TYPE "UDT_Divert_Constraint_Setting"
VERSION : 0.1
   STRUCT
      Enable : Bool := FALSE;
      Threshold : Int;
      Priority : Int;
      Sort_Code : Int;
      Preferred_Direction : Byte := 16#00;   // Bit0 = Wait Bit1= Straight Bit2= Left Bit3 = Right
      Disallowed_Direction : Byte := 16#00;   // Bit0 = Wait Bit1= Straight Bit2= Left Bit3 = Right
   END_STRUCT;

END_TYPE

TYPE "UDT_SWS_Servo_Setting"
VERSION : 0.1
   STRUCT
      Enable_Soft_Limit { ExternalAccessible := 'False'; ExternalVisible := 'False'; ExternalWritable := 'False'} : Bool := TRUE;
      Enable_Hard_Limit { ExternalAccessible := 'False'; ExternalVisible := 'False'; ExternalWritable := 'False'} : Bool;
      Continuous_Action_Mode : Bool := TRUE;
      STOUsed : Bool;
      Left_Position_Setpoint : Int := -60;   // [°]
      Right_Position_Setpoint : Int := 60;   // [°]
      Speed_Setpoint : Int := 1200;   // [°/s]
      Acc_Setpoint { ExternalAccessible := 'False'; ExternalVisible := 'False'; ExternalWritable := 'False'} : Int := 20000;   // [°/s²]
      Dec_Setpoint { ExternalAccessible := 'False'; ExternalVisible := 'False'; ExternalWritable := 'False'} : Int := 20000;   // [°/s²]
      Max_Left_Position { ExternalAccessible := 'False'; ExternalVisible := 'False'; ExternalWritable := 'False'} : Int := -65;   // [°]
      Max_Right_Position { ExternalAccessible := 'False'; ExternalVisible := 'False'; ExternalWritable := 'False'} : Int := 65;   // [°]
      Max_Speed { ExternalAccessible := 'False'; ExternalVisible := 'False'; ExternalWritable := 'False'} : Int := 1500;   // [°/s]
   END_STRUCT;

END_TYPE

TYPE "UDT_SWS_Roller_Hardware_Setting"
VERSION : 0.1
   STRUCT
      Module_Roller_Count : Int := 29;
      Speed_Straight : Int := 1200;
      Speed_Left : Int := 1500;
      Speed_Right : Int := 1500;
      Reference_RPM : Real := 470.0;
      Acceleration : Int := 4000;   // [mm/s²] Ramp up
      Deceleration : Int := 4000;   // [mm/s²] Ramp down
   END_STRUCT;

END_TYPE

TYPE "i_udtSettings"
VERSION : 0.1
   STRUCT
      timStartReadDelay : UDInt := 40;   // Start read delay time (mseconds)
      timSpare_Timer2 : UDInt;   // Not in use
      timNoActivity : UDInt := 10000;   // Time to consider Camera not working ok
      timTimeOutRead : UDInt := 400;   // TimeOut to get Barcode (mseconds)
      TimeStarting : UDInt := 5000;   // Time starting camera (waitting for normal operation)
      timTrshNoReadRow : Int;   // threshold no reads in a row
      xIndexProtocol : Bool := TRUE;   // 1: In Use; 0: Not used
      xIOConditioning : Bool := FALSE;   // 1: In Use; 0: Not used
      xFocusingDevice : Bool := FALSE;
      Protocol : Struct
         Encapsulation : Bool := TRUE;
         Header : String := '$02';
         Footer : String := '$03';
         Separator : String := '€';
         VirtualID : String := '!';
         ValidTelegram : String := '*';
         NoRead : String := '??????????';
         MultiRead : String := '9999999999';
      END_STRUCT;
      Telegrams : Struct
         Number : Int := 4;
         Parameters : Array[0..10] of Struct
            Length : Int;   // Telegram length without encapsulation
            "Type" : Int;   // 0: No Code; 1: Status Telegram; 2: Barcode Telegram; 9: Special Barcode Telegram
            ID : Char;   // Telegram ID. D: Status; I: Index Barcode
            Barcode : Struct   // Only for Types > 2
               FromDAD : String;
               ToPLC : String := '0000000000';
            END_STRUCT;
         END_STRUCT;
      END_STRUCT;
   END_STRUCT;

END_TYPE

TYPE "UDT_G115D_Setting"
VERSION : 0.1
   STRUCT
      Speed1 : Int := 1000;   // [mm/s] Target speed 1
      Speed2 : Int := 500;   // [mm/s] Target speed 2
      Speed3 : Int;   // [mm/s] Target speed 3
      Speed4 : Int;   // [mm/s] Target speed 4
      Acceleration : Int := 4000;   // [mm/s²] Ramp up
      Deceleration : Int := 4000;   // [mm/s²] Ramp down
      RefSpeed : Int;   // [mm/s] Speed at 3000RPM
      RefRampTime : Int := 10000;   // [ms] Ramp up and ramp down time for 3000RPM
      Magnetization_Delay : Int;   // [ms] Delay time from run command to mote have speed
      ReverseDirection : Bool;   // TRUE = Reverse inverter output direction
      STOUsed : Bool;   // TRUE = STO is used
   END_STRUCT;

END_TYPE

TYPE "UDT_MultiControl_HW_Diagnostics"
VERSION : 0.1
   STRUCT
      RD1_Run_Command : Bool;   // Rum command from controller
      RD2_Run_Command : Bool;   // Rum command from controller
      RD3_Run_Command : Bool;   // Rum command from controller
      RD4_Run_Command : Bool;   // Rum command from controller
      RD1_Actual_Speed : Int;   // [mm/s] Motor actual speed
      RD2_Actual_Speed : Int;   // [mm/s] Motor actual speed
      RD3_Actual_Speed : Int;   // [mm/s] Motor actual speed
      RD4_Actual_Speed : Int;   // [mm/s] Motor actual speed
      Control_Voltage : Int;   // [mV] Control logic voltage
      Motor_Voltage : Int;   // [mV] Motor voltage
      Temperature : Int;   // [0,1°] Temperature
      RD1_Actual_Current : Int;   // [mA] Actual current
      RD2_Actual_Current : Int;   // [mA] Actual current
      RD3_Actual_Current : Int;   // [mA] Actual current
      RD4_Actual_Current : Int;   // [mA] Actual current
      Motor_Start_Stop_Count : UInt;   // Count of motor start and stop
      Motor_Direction_Switch_Count : UInt;   // Count of motor switch direction
      Motor_Started_Time : UDInt;   // [s] Count time of motor running
   END_STRUCT;

END_TYPE

TYPE "UDT_PEC_Position_Setting"
TITLE = UDT_Sett_PEC
VERSION : 0.1
//Setting of photo electric cell
//# Block Info
//- Title:            UDT_Sett_PEC
//- Comment/Function: Setting of photo electric cell
//- Library/Family:   APS
//- Author:           Jay Liu
//- Tested with:      ---
//- Engineering:      TIA Portal V20
//- Restrictions:     ---
//- Requirements:     ---
//
//# History
// |Version  | Date       | Author                 | Description                   |
// |---------|------------|------------------------|------------------------------ |
// |01.00.00 | 2026-01-22 | Jay Liu                | First released version        |
   STRUCT
      Blockage_Length : DInt := 3000;   // [mm] Delay for detecting a PEC blockage during the running
      Delay_On : DInt := 50;   // [mm] Delay on leading edge of product (flap filter)
      Delay_Off : DInt := 50;   // [mm] Delay off trailing edge of product (flap filter)
      Shifting_Offset : DInt;   // [mm] Shift offset of PE signal
      Handover_Offset : DInt;   // [mm] Distance between PE and the end of section
      Detect_PEC_OnStopped : Bool := TRUE;   // TRUE = Enable delay timer even the section is not running
      Reset_Block_PEC_Oc : Bool;   // TRUE = Allow reset of blockage error with PEC still covered
      Item_On : Bool;   // TRUE = When detect item the input signal should be true FALSE= When detect item the input signal should be false
   END_STRUCT;

END_TYPE

TYPE "UDT_TCON_PAR"
VERSION : 0.1
   STRUCT
      InterfaceId : HW_ANY := 64;
      ID : CONN_OUC := 1;
      ConnectionType : Byte := 11;
      ActiveEstablished : Bool;
      RemoteAddress {InstructionName := 'IP_V4'; LibVersion := '1.0'} : IP_V4;
      RemotePort : UInt;
      LocalPort : UInt := 6000;
   END_STRUCT;

END_TYPE

TYPE "UDT_Divert_Decision_Setting"
VERSION : 0.1
   STRUCT
      Decision_Position : DInt;
      Straight_Destination { S7_SetPoint := 'True'} : Int;
      Left_Destination { S7_SetPoint := 'True'} : Int;
      Right_Destination { S7_SetPoint := 'True'} : Int;
      High_Priority { S7_SetPoint := 'True'} : Int := 2;   // Bit0 = Wait Bit1= Straight Bit2= Left Bit3 = Right
      Middle_Priority { S7_SetPoint := 'True'} : Int := 4;   // Bit0 = Wait Bit1= Straight Bit2= Left Bit3 = Right
      Low_Priority { S7_SetPoint := 'True'} : Int := 8;   // Bit0 = Wait Bit1= Straight Bit2= Left Bit3 = Right
      Default_Direction : Int := 8;   // Bit0 = Wait Bit1= Straight Bit2= Left Bit3 = Right
      Allow_Wait : Bool := FALSE;
      Destination_Invalid : "UDT_Divert_Constraint_Setting" := ((), (), 1, 7, (), ());
      No_Destination : "UDT_Divert_Constraint_Setting" := ((), (), 2, 16, (), ());
      Gap_Error : "UDT_Divert_Constraint_Setting" := ((), 250, 4, 4, (), ());
      Diemension_Error : "UDT_Divert_Constraint_Setting" := ((), 700, 6, 18, (), ());
      Throughput_Limit_Straight : "UDT_Divert_Constraint_Setting" := ((), (), 10, 13, (), ());
      Throughput_Limit_Left : "UDT_Divert_Constraint_Setting" := ((), (), 10, 13, (), ());
      Throughput_Limit_Right : "UDT_Divert_Constraint_Setting" := ((), (), 10, 13, (), ());
      Dir_Fault_Straight : "UDT_Divert_Constraint_Setting" := ((), (), 13, 20, (), ());
      Dir_Fault_Left : "UDT_Divert_Constraint_Setting" := ((), (), 13, 20, (), ());
      Dir_Fault_Right : "UDT_Divert_Constraint_Setting" := ((), (), 13, 20, (), ());
      Dir_Disabled_Straight : "UDT_Divert_Constraint_Setting" := ((), (), 14, 12, (), ());
      Dir_Disabled_Left : "UDT_Divert_Constraint_Setting" := ((), (), 14, 12, (), ());
      Dir_Disabled_Right : "UDT_Divert_Constraint_Setting" := ((), (), 14, 12, (), ());
      Dir_Full_Straight : "UDT_Divert_Constraint_Setting" := ((), (), 15, 5, (), ());
      Dir_Full_Left : "UDT_Divert_Constraint_Setting" := ((), (), 15, 5, (), ());
      Dir_Full_Right : "UDT_Divert_Constraint_Setting" := ((), (), 15, 5, (), ());
      No_Read : "UDT_Divert_Constraint_Setting" := ((), (), 16, 8, (), ());
      No_Code : "UDT_Divert_Constraint_Setting" := ((), (), 17, 9, (), ());
      Multi_Read : "UDT_Divert_Constraint_Setting" := ((), (), 18, 10, (), ());
      Unexpected_Item : "UDT_Divert_Constraint_Setting" := ((), (), 19, 2, (), ());
   END_STRUCT;

END_TYPE

TYPE "UDT_SWS_Divert_Setting"
VERSION : 0.1
   STRUCT
      Fixed_Ratio_Staight : Int;
      Fixed_Ratio_Left : Int;
      Fixed_Ratio_Right : Int;
      First_Group_Action_Delay : Int := 350;
      Group2_Action_Delay : Int := 160;
      Group3_Action_Delay : Int := 160;
      Group4_Action_Delay : Int := 160;
      Group5_Action_Delay : Int := 160;
      Group6_Action_Delay : Int := 160;
      Group7_Action_Delay : Int := 160;
      Group8_Action_Delay : Int := 160;
      Group9_Action_Delay : Int := 160;
   END_STRUCT;

END_TYPE

TYPE "UDT_SWS_Hardware_Setting"
VERSION : 0.1
   STRUCT
      Roller { S7_SetPoint := 'False'} : "UDT_SWS_Roller_Hardware_Setting" := (29, 1200, 1500, 1500, 470.0, 4000, 4000);
      Servo_U401 : "UDT_SWS_Servo_Setting" := ((), (), (), (), -30, 30, (), (), (), (), (), ());
      Servo_U411 : "UDT_SWS_Servo_Setting" := ((), (), (), (), -45, 45, (), (), (), (), (), ());
      Servo_U421 : "UDT_SWS_Servo_Setting";
      Servo_U431 : "UDT_SWS_Servo_Setting";
      Servo_U441 : "UDT_SWS_Servo_Setting";
      Servo_U451 : "UDT_SWS_Servo_Setting";
      Servo_U461 : "UDT_SWS_Servo_Setting";
      Servo_U471 : "UDT_SWS_Servo_Setting";
      Servo_U481 : "UDT_SWS_Servo_Setting";
   END_STRUCT;

END_TYPE

TYPE "UDT_MultiControl_Setting"
VERSION : 0.1
   STRUCT
      Speed1 : Int := 1000;   // [mm/s] Target speed 1
      Speed2 : Int := 500;   // [mm/s] Target speed 2
      Speed3 : Int;   // [mm/s] Target speed 3
      Speed4 : Int;   // [mm/s] Target speed 4
      Acceleration : Int := 4000;   // [mm/s²] Ramp up
      Deceleration : Int := 4000;   // [mm/s²] Ramp down
      RefSpeed : Int := 1390;   // [mm/s] Reference Speed
      RD1_Motor_Number : Int;
      RD2_Motor_Number : Int;
      RD3_Motor_Number : Int;
      RD4_Motor_Number : Int;
      ReverseDirection : Bool;
   END_STRUCT;

END_TYPE

TYPE "UDT_G115D_HW_Diagnostics"
VERSION : 0.1
   STRUCT
      Run_Command : Bool;   // Rum command from controller
      Brake_Open : Bool;   // Holding brake open
      DI0 : Bool;   // Digital input 0 status
      DI1 : Bool;   // Digital input 1 status
      DI2 : Bool;   // Digital input 2 status
      DI3 : Bool;   // Digital input 3 status
      DIO24 : Bool;   // Digital input/output 24 status
      DIO25 : Bool;   // Digital input/output 25 status
      Memory_Card_In : Bool;   // Memory card is inserted
      Memory_Card_Active : Bool;   // Memory card is active
      PN_Port1_Down : Bool;   // Profinet port 1 up
      PN_Port2_Down : Bool;   // Profinet port 2 up
      Actual_Speed : Int;   // [mm/s] Motor Actual Speed
      DCLink_Voltage : Int;   // [V] DC link voltage
      Actual_Current : Int;   // [0.1A] Actual current
      Active_Power : Int;   // [W] Active power
      Motor_Start_Stop_Count : UInt;   // Count of motor start and stop
      Motor_Direction_Switch_Count : UInt;   // Count of motor switch direction
      Motor_Started_Time : UDInt;   // [s] Count time of motor running
   END_STRUCT;

END_TYPE

TYPE "UDT_SWS_Roller_Interface_Setting"
VERSION : 0.1
   STRUCT
      Status_Interval : Time := T#200ms;
      Num_Of_Comm_Error : Int := 3;
   END_STRUCT;

END_TYPE

TYPE "UDT_G115D_HW_Input"
VERSION : 0.1
   STRUCT
      ZSW1_Bit00_ReadyOn : Bool;   // 0: Ready for switching on
      ZSW1_Bit01_Ready : Bool;   // 1: Ready (operating condition)
      ZSW1_Bit02_Enabled : Bool;   // 2: Operation enabled
      ZSW1_Bit03_Fault : Bool;   // 3: Fault present (1: fault)
      ZSW1_Bit04_NoCoastActive : Bool;   // 4: No coast down active (0: active)
      ZSW1_Bit05_NoQuickStopActive : Bool;   // 5: No quick stop active (0: active)
      ZSW1_Bit06_Inhibit : Bool;   // 6: Switching on inhibited
      ZSW1_Bit07_Alarm : Bool;   // 7: Alarm present (1: alarm)
      ZSW1_Bit08_DeviationOK : Bool;   // 8: Setpoint/actual value deviation
      ZSW1_Bit09_ControlQuest : Bool;   // 9: Control requested
      ZSW1_Bit10_OverSpeed : Bool;   // 10: f or n comparison value reached
      ZSW1_Bit11_Limit : Bool;   // 11: Torque limit not reached
      ZSW1_Bit12_Brake : Bool;   // 12: Holding brake open
      ZSW1_Bit13_MotorTempOK : Bool;   // 13: Motor temperature OK (1: OK)
      ZSW1_Bit14_Direction_CW : Bool;   // 14: n_act >= 0 (1: positive)
      ZSW1_Bit15_VFDTempOK : Bool;   // 15: Reserved Speed actual value (NIST_A)
      NIST_A : Int;   // Actual speed (-16384 to +16384)
      ZSW_G115D_Bit00_DI0 : Bool;   // 0: Digital input 0 status
      ZSW_G115D_Bit01_DI1 : Bool;   // 1: Digital input 1 status
      ZSW_G115D_Bit02_DI2 : Bool;   // 2: Digital input 2 status
      ZSW_G115D_Bit03_DI3 : Bool;   // 3: Digital input 3 status
      ZSW_G115D_Bit04_DIO24 : Bool;   // 4: DI/O 24 status
      ZSW_G115D_Bit05_DIO25 : Bool;   // 5: DI/O 25 status
      ZSW_G115D_Bit06_STOActive : Bool;   // 6: STO is active
      ZSW_G115D_Bit07_Reserved : Bool;   // 7: Reserved
      ZSW_G115D_Bit08_PowerOff : Bool;   // 8: Power switch OFF status
      ZSW_G115D_Bit09_Auto : Bool;   // 9: Automatic mode active
      ZSW_G115D_Bit10_Manual : Bool;   // 10: Manual mode active
      ZSW_G115D_Bit11_Bypass : Bool;   // 11: Stop/Slow bypass activated
      ZSW_G115D_Bit12_ContMotion : Bool;   // 12: Continuous motion activated
      ZSW_G115D_Bit13_JogLeft : Bool;   // 13: Motor jogging to the left
      ZSW_G115D_Bit14_JogRight : Bool;   // 14: Motor jogging to the right
      ZSW_G115D_Bit15_Reserved : Bool;   // 15: Reserved Fault and alarm codes
      FaultCode : Word;   // Fault code (0: no fault)
      AlarmCode : Word;   // Alarm code (0: no alarm)
      DCLinkVoltage : Int;   // DC link voltage [V]
      ActualCurrent : Int;   // Actual current [0.1A]
      ActivePower : Int;   // Active power [W]
      ZSW2_G115D_Bit00_Memory_Card_In : Bool;
      ZSW2_G115D_Bit01_Memory_Card_Active : Bool;
      ZSW2_G115D_Bit02_Memory_Card_Siemens : Bool;
      ZSW2_G115D_Bit03_Memory_Card_USB : Bool;
      ZSW2_G115D_Bit04_Reserved : Bool;
      ZSW2_G115D_Bit05_Reserved : Bool;
      ZSW2_G115D_Bit06_Reserved : Bool;
      ZSW2_G115D_Bit07_Reserved : Bool;
      ZSW2_G115D_Bit08_Reserved : Bool;
      ZSW2_G115D_Bit09_Reserved : Bool;
      ZSW2_G115D_Bit10_Reserved : Bool;
      ZSW2_G115D_Bit11_Reserved : Bool;
      ZSW2_G115D_Bit12_Reserved : Bool;
      ZSW2_G115D_Bit13_Reserved : Bool;
      ZSW2_G115D_Bit14_Reserved : Bool;
      ZSW2_G115D_Bit15_Reserved : Bool;
   END_STRUCT;

END_TYPE

TYPE "UDT_S210_Speed_Setting"
VERSION : 0.1
   STRUCT
      Speed1 : Int := 1000;   // [mm/s] Target speed 1
      Speed2 : Int := 500;   // [mm/s] Target speed 2
      Speed3 : Int;   // [mm/s] Target speed 3
      Speed4 : Int;   // [mm/s] Target speed 4
      Acceleration : Int := 4000;   // [mm/s²] Ramp up
      Deceleration : Int := 4000;   // [mm/s²] Ramp down
      MinSpeed : Int := 500;   // [mm/s] Minimum target speed
      MaxSpeed : Int := 2500;   // [mm/s] Maximum target speed
      Continuous_Action_Mode : Bool := TRUE;
      Use_Hardware_Feedback : Bool;
      ReverseDirection : Bool;
      STOUsed : Bool;
   END_STRUCT;

END_TYPE

TYPE "UDT_G115D_HW_Output"
VERSION : 0.1
   STRUCT
      STW1_Bit00_On : Bool;   // 0: ON/OFF1 command (0->1: ON)
      STW1_Bit01_Off2 : Bool;   // 1: No OFF2 command (0: active, coast stop)
      STW1_Bit02_Off3 : Bool;   // 2: No OFF3 command (0: active, quick stop)
      STW1_Bit03_Enable : Bool;   // 3: Operation enable
      STW1_Bit04_RampEnable : Bool;   // 4: Ramp-function generator enable
      STW1_Bit05_RampContinue : Bool;   // 5: Continue ramp-function generator
      STW1_Bit06_SetEnable : Bool;   // 6: Setpoint enable
      STW1_Bit07_Ack : Bool;   // 7: Acknowledge faults (0->1: acknowledge)
      STW1_Bit08_Reserved : Bool;   // 8: Reserved
      STW1_Bit09_Reserved : Bool;   // 9: Reserved
      STW1_Bit10_PLC : Bool;   // 10: Control by PLC (must be 1)
      STW1_Bit11_Reverse : Bool;   // 11: Reverse (1: reverse direction)
      STW1_Bit12_Reserved : Bool;   // 12: Reserved
      STW1_Bit13_MOP_Up : Bool;   // 13: Motorized potentiometer, raise
      STW1_Bit14_MOP_Down : Bool;   // 14: Motorized potentiometer, lower
      STW1_Bit15_Reserved : Bool;   // 15: Reserved Speed setpoint (NSOLL_A)
      NSOLL_A : Int;   // Speed setpoint (-16384 to +16384)
      STW_G115D_Bit00_DO24 : Bool;   // 0: DO 24 control
      STW_G115D_Bit01_DO25 : Bool;   // 1: DO 25 control
      STW_G115D_Bit02_Disable_StopSlow_Sensor : Bool;   // 2: Stop-Slow bypass
      STW_G115D_Bit03_Reserved : Bool;   // 3: Reserved
      STW_G115D_Bit04_Reserved : Bool;   // 4: Reserved
      STW_G115D_Bit05_Reserved : Bool;   // 5: Reserved
      STW_G115D_Bit06_Reserved : Bool;   // 6: Reserved
      STW_G115D_Bit07_Reserved : Bool;   // 7: Reserved
      STW_G115D_Bit08_Reserved : Bool;   // 8: Reserved
      STW_G115D_Bit09_Reserved : Bool;   // 9: Reserved
      STW_G115D_Bit10_Reserved : Bool;   // 10: Reserved
      STW_G115D_Bit11_Reserved : Bool;   // 11: Reserved
      STW_G115D_Bit12_Reserved : Bool;   // 12: Reserved
      STW_G115D_Bit13_Reserved : Bool;   // 13: Reserved
      STW_G115D_Bit14_Reserved : Bool;   // 14: Reserved
      STW_G115D_Bit15_Reserved : Bool;   // 15: Reserved
      RampUpScaling : Int;   // Ramp-up time scaling (0-200% = 0-32767)
      RampDownScaling : Int;   // Ramp-down time scaling (0-200% = 0-32767)
   END_STRUCT;

END_TYPE

TYPE "UDT_S210_HW_Diagnostics"
VERSION : 0.1
   STRUCT
      Run_Command : Bool;   // Rum command from controller
      DI0 : Bool;   // Digital input 0 status
      DI1 : Bool;   // Digital input 1 status
      DI2 : Bool;   // Digital input 2 status
      DI3 : Bool;   // Digital input 3 status
      DI4 : Bool;   // Digital input 4 status
      PN_Port1_Down : Bool;   // Profinet port 1 up
      PN_Port2_Down : Bool;   // Profinet port 2 up
      Actual_Speed : Int;   // [mm/s] Motor actual speed
      Actual_Displacement : Int;   // [mm/scan] Motor movement distance
      Actual_Position : Real;   // [°] Motor actual position
      DCLink_Voltage : Int;   // [V] DC link voltage
      Actual_Current : Int;   // [0.1A] Actual current
      Active_Power : Int;   // [W] Active power
      Motor_Start_Stop_Count : UInt;   // Count of motor start and stop
      Motor_Direction_Switch_Count : UInt;   // Count of motor switch direction
      Motor_Started_Time : UDInt;   // [s] Count time of motor running
   END_STRUCT;

END_TYPE

TYPE "UDT_Base_Conveyor_Setting"
TITLE = UDT_Sett_Base_Conveyor
VERSION : 0.1
//Setting of base tranpsort control
//# Block Info
//- Title:            UDT_Sett_Base_Conveyor
//- Comment/Function: Setting of base tranpsort control
//- Library/Family:   APS
//- Author:           Jay Liu
//- Tested with:      ---
//- Engineering:      TIA Portal V20
//- Restrictions:     ---
//- Requirements:     ---
//
//# History
// |Version  | Date       | Author                 | Description                   |
// |---------|------------|------------------------|------------------------------ |
// |01.00.00 | 2026-01-22 | Jay Liu                | First released version        |
   STRUCT
      Delay_Dieback : DInt := 50;   // [mm] Delay from end to stop in dieback
      Delay_Startup : DInt := 100;   // [mm] Delay restart after dieback
      Delay_Waiting_Item : DInt;   // [mm] Delay for receive item from upstream
      Delay_Finish_Handover : DInt;   // [mm] Delay handover after items exit the END PEC
      Delay_Energysave : DInt := 5000;   // [mm] Delay running after clearing
      Delay_Cascade_Startup : DInt := 100;   // [mm] Cascade delay 0: Startup immediately
      Delay_Cascade_Shutdown : DInt := -1;   // [ms] Cascade delay -1: disable function 0: Shutdown immediately
      Slave_Mode : Bool;   // TRUE = Make this section a slave
      Enable_DieForward : Bool;   // TRUE = Halt conveyor if upstream handover occurs error
   END_STRUCT;

END_TYPE

TYPE "UDT_Flow_Control_Setting"
TITLE = UDT_Sett_Flow_Control
VERSION : 0.1
//Setting of flow control
//# Block Info
//- Title:            UDT_Sett_Flow_Control
//- Comment/Function: Setting of flow control
//- Library/Family:   APS
//- Author:           Jay Liu
//- Tested with:      ---
//- Engineering:      TIA Portal V20
//- Restrictions:     ---
//- Requirements:     ---
//
//# History
// |Version  | Date       | Author                 | Description                   |
// |---------|------------|------------------------|------------------------------ |
// |01.00.00 | 2026-01-22 | Jay Liu                | First released version        |
   STRUCT
      Minimum_Gap : Int;   // [mm] Minimum gap length between products (0 = no gap control)
      Add_Gap_Stop : Int;   // [mm] Additional gap after stop of upstream conveyor
      Minimum_Head_To_Head : Int;   // [mm] Minimum head to head length (0 = no head to head control)
      Add_Head_To_Head_Stop : Int;   // [mm] Additional head to head length after stop of upstream conveyor
   END_STRUCT;

END_TYPE

TYPE "UDT_PEC_Trigger_Setting"
TITLE = UDT_Sett_PEC
VERSION : 0.1
//Setting of photo electric cell
//# Block Info
//- Title:            UDT_Sett_PEC
//- Comment/Function: Setting of photo electric cell
//- Library/Family:   APS
//- Author:           Jay Liu
//- Tested with:      ---
//- Engineering:      TIA Portal V20
//- Restrictions:     ---
//- Requirements:     ---
//
//# History
// |Version  | Date       | Author                 | Description                   |
// |---------|------------|------------------------|------------------------------ |
// |01.00.00 | 2026-01-22 | Jay Liu                | First released version        |
   STRUCT
      Blockage_Length : Int := 3000;   // [mm] Delay for detecting a PEC blockage during the running
      Delay_On : Int := 50;   // [mm] Delay on leading edge of product (flap filter)
      Delay_Off : Int := 50;   // [mm] Delay off trailing edge of product (flap filter)
      Detect_PEC_OnStopped : Bool := TRUE;   // TRUE = Enable delay timer even the section is not running
      Reset_Block_PEC_Oc : Bool;   // TRUE = Allow reset of blockage error with PEC still covered
      Item_On : Bool;   // TRUE = When detect item the input signal should be true FALSE= When detect item the input signal should be false
   END_STRUCT;

END_TYPE

TYPE "UDT_Track_Statistics"
VERSION : 0.1
   STRUCT
      Last_Slip : Int;
      Last_Data : Int;
      Average_Slip : Real;
      Update_Performance : Real;
      Missing_Items : UDInt;
      UFO_Generated : UDInt;
      Number_Of_Items : UDInt;
   END_STRUCT;

END_TYPE

TYPE "UDT_Mesasuring_Point_Statistics"
VERSION : 0.1
   STRUCT
      Capacity : Int;
      Length : UDInt;
      Window : UDInt;
      Gap : UDInt;
   END_STRUCT;

END_TYPE

TYPE "UDT_Scanner_Statistics"
VERSION : 0.1
   STRUCT
      Total : UDInt;
      GoodRead : UDInt;
      NoRead : UDInt;
      MultiRead : UDInt;
      NoCode : UDInt;
      NoFoundID : UDInt;
      NotDefined : UDInt;
   END_STRUCT;

END_TYPE

TYPE "UDT_Chute_Statistics"
VERSION : 0.1
   STRUCT
      PE_Full_Items : UDInt;
   END_STRUCT;

END_TYPE

TYPE "UDT_IODevice_Diag"
TITLE = UDT_Diag_HW
VERSION : 0.1
//Diagnose data of IO Device
//# Block Info
//- Title:            UDT_Diag_HW
//- Comment/Function: Diagnose data of IO Device
//- Library/Family:   APS
//- Author:           Jay Liu
//- Tested with:      ---
//- Engineering:      TIA Portal V20
//- Restrictions:     ---
//- Requirements:     ---
//
//# History
// |Version  | Date       | Author                 | Description                   |
// |---------|------------|------------------------|------------------------------ |
// |01.00.00 | 2026-01-22 | Jay Liu                | First released version        |
   STRUCT
      Module_Not_Present : Array[0..127] of Bool;   // Module not present
      Module_Error : Array[0..127] of Bool;   // Module error
   END_STRUCT;

END_TYPE

TYPE "UDT_PNIO_System_Diag"
TITLE = UDT_Diag_PNIO_System
VERSION : 0.1
//Diagnose data of IO System
//# Block Info
//- Title:            UDT_Diag_PNIO_System
//- Comment/Function: Diagnose data of IO System
//- Library/Family:   APS
//- Author:           Jay Liu
//- Tested with:      ---
//- Engineering:      TIA Portal V20
//- Restrictions:     ---
//- Requirements:     ---
//
//# History
// |Version  | Date       | Author                 | Description                   |
// |---------|------------|------------------------|------------------------------ |
// |01.00.00 | 2026-01-22 | Jay Liu                | First released version        |
   STRUCT
      Device_Not_Present : Array[0..1023] of Bool;   // Profinet device not present
      Device_Error : Array[0..1023] of Bool;   // Profinet device error
   END_STRUCT;

END_TYPE

TYPE "UDT_Divert_Statistics"
VERSION : 0.1
   STRUCT
      Direction_Straight : UDInt;
      Direction_Left : UDInt;
      Direction_Right : UDInt;
   END_STRUCT;

END_TYPE

TYPE "UDT_G115D_HW_Interface"
VERSION : 0.1
   STRUCT
      Input { S7_SetPoint := 'False'} : "UDT_G115D_HW_Input";
      Output : "UDT_G115D_HW_Output";
   END_STRUCT;

END_TYPE

TYPE "UDT_Conv_Multiple_S210_Diagnostics"
VERSION : 0.1
   STRUCT
      RTS : Bool;   // Section ready to send item
      TIP : Bool;   // Section transfer in porgress
      Downstream_RTR : Bool;   // Downstream section ready to receive item
      Items_Count : UDInt;   // Count of items passed
      Displacement : Int;   // [mm/scan] Conveyor movement distance
      Hardware_U01 { S7_SetPoint := 'False'} : "UDT_S210_HW_Diagnostics";
      Hardware_U02 : "UDT_S210_HW_Diagnostics";
      Hardware_U03 : "UDT_S210_HW_Diagnostics";
      Hardware_U04 : "UDT_S210_HW_Diagnostics";
      Hardware_U05 : "UDT_S210_HW_Diagnostics";
      Hardware_U06 : "UDT_S210_HW_Diagnostics";
      Hardware_U07 : "UDT_S210_HW_Diagnostics";
      Hardware_U08 : "UDT_S210_HW_Diagnostics";
      Hardware_U09 : "UDT_S210_HW_Diagnostics";
      Hardware_U10 : "UDT_S210_HW_Diagnostics";
   END_STRUCT;

END_TYPE

TYPE "UDT_Conv_Dual_G115D_Diagnostics"
VERSION : 0.1
   STRUCT
      RTS : Bool;   // Section ready to send item
      TIP : Bool;   // Section transfer in porgress
      Downstream_RTR : Bool;   // Downstream section ready to receive item
      Items_Count : UDInt;   // Count of items passed
      Displacement : Int;   // [mm/scan] Conveyor movement distance
      Hardware_U01 { S7_SetPoint := 'False'} : "UDT_G115D_HW_Diagnostics";   // Invert driver
      Hardware_U02 : "UDT_G115D_HW_Diagnostics";
   END_STRUCT;

END_TYPE

TYPE "UDT_Conv_Triple_G115D_Diagnostics"
VERSION : 0.1
   STRUCT
      RTS : Bool;   // Section ready to send item
      TIP : Bool;   // Section transfer in porgress
      Downstream_RTR : Bool;   // Downstream section ready to receive item
      Items_Count : UDInt;   // Count of items passed
      Displacement : Int;   // [mm/scan] Conveyor movement distance
      Hardware_U01 { S7_SetPoint := 'False'} : "UDT_G115D_HW_Diagnostics";   // Invert driver
      Hardware_U02 : "UDT_G115D_HW_Diagnostics";
      Hardware_U03 : "UDT_G115D_HW_Diagnostics";
   END_STRUCT;

END_TYPE

TYPE "UDT_Conv_MultiControl_Diagnostics"
VERSION : 0.1
   STRUCT
      RTS : Bool;   // Section ready to send item
      TIP : Bool;   // Section transfer in porgress
      Downstream_RTR : Bool;   // Downstream section ready to receive item
      Items_Count : UDInt;   // Count of items passed
      Displacement : Int;   // [mm/scan] Conveyor movement distance
      Hardware_U01 { S7_SetPoint := 'False'} : "UDT_MultiControl_HW_Diagnostics";   // Invert driver
      Hardware_U02 : "UDT_MultiControl_HW_Diagnostics";
      Hardware_U03 : "UDT_MultiControl_HW_Diagnostics";
      Hardware_U04 : "UDT_MultiControl_HW_Diagnostics";
   END_STRUCT;

END_TYPE

TYPE "UDT_Conv_G115D_Diagnostics"
VERSION : 0.1
   STRUCT
      RTS : Bool;   // Section ready to send item
      TIP : Bool;   // Section transfer in porgress
      Downstream_RTR : Bool;   // Downstream section ready to receive item
      Items_Count : UDInt;   // Count of items passed
      Displacement : Int;   // [mm/scan] Conveyor movement distance
      Hardware { S7_SetPoint := 'False'} : "UDT_G115D_HW_Diagnostics";   // Invert driver
   END_STRUCT;

END_TYPE

TYPE "UDT_MultiControl_HW_Input"
VERSION : 0.1
   STRUCT
      Sensor1 : Bool;
      Sensor2 : Bool;
      Sensor3 : Bool;
      Sensor4 : Bool;
      Sensor5 : Bool;
      Sensor6 : Bool;
      Sensor7 : Bool;
      Sensor8 : Bool;
      Digital_Input_1 : Bool;
      Digital_Input_2 : Bool;
      Digital_Input_3 : Bool;
      Digital_Input_4 : Bool;
      Digital_Input_Spare_1 : Bool;
      Digital_Input_Spare_2 : Bool;
      Digital_Input_Spare_3 : Bool;
      Digital_Input_Spare_4 : Bool;
      MotorErr_RD1 : Bool;
      MotorErr_RD2 : Bool;
      MotorErr_RD3 : Bool;
      MotorErr_RD4 : Bool;
      MotorSpeed_RD1 : SInt;
      MotorSpeed_RD2 : SInt;
      MotorSpeed_RD3 : SInt;
      MotorSpeed_RD4 : SInt;
      MotorStates_Spare : Byte;
      MotorCurrent_RD1 : Int;   // [mA]
      MotorCurrent_RD2 : Int;   // [mA]
      MotorCurrent_RD3 : Int;   // [mA]
      MotorCurrent_RD4 : Int;   // [mA]
      Voltage_Motor : Int;   // [mV]
      Voltage_Control : Int;   // [mV]
      Temperature : Int;   // [0.1C]
      SystemUpTime : UDInt;   // [s]
   END_STRUCT;

END_TYPE

TYPE "UDT_Merge_Singulator_Setting"
VERSION : 0.1
   STRUCT
      StartUp_Delay : Int;   // [ms]
      Dieback_Delay : Int;   // [ms]
   END_STRUCT;

END_TYPE

TYPE "UDT_Echelon_Setting"
VERSION : 0.1
   STRUCT
      StartUp_Delay : Int;   // [ms]
      Dieback_Delay : Int;   // [ms]
   END_STRUCT;

END_TYPE

TYPE "UDT_Tipper_Setting"
VERSION : 0.1
   STRUCT
      StartUp_Delay : Int;   // [ms]
      Dieback_Delay : Int;   // [ms]
   END_STRUCT;

END_TYPE

TYPE "UDT_Datalogic_AV900_Setting"
VERSION : 0.1
   STRUCT
      Trigger_Position : DInt;
      Scanner_ID : String[16];
      Interface { S7_SetPoint := 'False'} : "i_udtSettings";
   END_STRUCT;

END_TYPE

TYPE "UDT_PLC_Log_Setting"
VERSION : 0.1
   STRUCT
      Minimum_Log_Level : Int := 3;   // 1: Trace 2: Debug 3: Info 4: Warn 5: Error 6: Fatal
      Connection { S7_SetPoint := 'False'} : "UDT_TCON_PAR";
   END_STRUCT;

END_TYPE

TYPE "UDT_AWCS_Setting"
VERSION : 0.1
   STRUCT
      InterfaceId : HW_ANY := 72;
      ID_Range : Int := 1;
      LocalPort : UInt := 3000;
   END_STRUCT;

END_TYPE

TYPE "UDT_SSM_Setting"
TITLE = UDT_Sett_SSM
VERSION : 0.1
//Setting of start stop manager
//# Block Info
//- Title:            UDT_Sett_SSM
//- Comment/Function: Setting of start stop manager
//- Library/Family:   APS
//- Author:           Jay Liu
//- Tested with:      ---
//- Engineering:      TIA Portal V20
//- Restrictions:     ---
//- Requirements:     ---
//
//# History
// |Version  | Date       | Author                 | Description                   |
// |---------|------------|------------------------|------------------------------ |
// |01.00.00 | 2026-01-22 | Jay Liu                | First released version        |
   STRUCT
      StartUp_Indication_Time : Int;   // [s] Duration of Start-Up indication
      Restart_Indication_Time : Int;   // [s] Duration of Restart indication
      ControlStop_Time : Int;   // [s] Time out on controlled stop
   END_STRUCT;

END_TYPE

TYPE "UDT_SWS_Roller_Module_Motor_Status"
VERSION : 0.1
   STRUCT
      None : Bool;
      NotConnected : Bool;
      Blockage : Bool;
      OK : Bool;
   END_STRUCT;

END_TYPE

TYPE "UDT_S210_HW_Output"
VERSION : 0.1
   STRUCT
      STW1_Bit00_On : Bool;   // 0: ON/OFF1 command (0->1: ON)
      STW1_Bit01_Off2 : Bool;   // 1: OFF2 command (0: active, coast stop)
      STW1_Bit02_Off3 : Bool;   // 2: OFF3 command (0: active, quick stop)
      STW1_Bit03_Enable : Bool;   // 3: Operation enable
      STW1_Bit04_NotRejectTask : Bool;   // 4: Not reject traversing task
      STW1_Bit05_NoIntermediateStop : Bool;   // 5: Intermediate stop (0: active)
      STW1_Bit06_ActivateTask : Bool;   // 6: Activate traversing task (0->1: start)
      STW1_Bit07_Ack : Bool;   // 7: Acknowledge faults (0->1: acknowledge)
      STW1_Bit08_Jog1 : Bool;   // 8: Jog 1 signal source
      STW1_Bit09_Jog2 : Bool;   // 9: Jog 2 signal source
      STW1_Bit10_PLC : Bool;   // 10: Control by PLC (must be 1)
      STW1_Bit11_StartHoming : Bool;   // 11: Start homing (0â†’1: start)
      STW1_Bit12_Reserved : Bool;   // 12: Reserved
      STW1_Bit13_ExtBlockChange : Bool;   // 13: External block change
      STW1_Bit14_Reserved : Bool;   // 14: Reserved
      STW1_Bit15_Reserved : Bool;   // 15: Reserved
      POS_STW1_Bit00_Traversing0 : Bool;   // 0: Traversing clock selection, bit 0
      POS_STW1_Bit01_Traversing1 : Bool;   // 1: Traversing clock selection, bit 1
      POS_STW1_Bit02_Traversing2 : Bool;   // 2: Traversing clock selection, bit 2
      POS_STW1_Bit03_Traversing3 : Bool;   // 3: Traversing clock selection, bit 3
      POS_STW1_Bit04_Traversing4 : Bool;   // 4: Traversing clock selection, bit 4
      POS_STW1_Bit05_Traversing5 : Bool;   // 5: Traversing clock selection, bit 5
      POS_STW1_Bit06_Reserved : Bool;   // 6: Reserved
      POS_STW1_Bit07_ReleaseBrake : Bool;   // 7: The converter opens a connected holding brake
      POS_STW1_Bit08_Absolute : Bool;   // 8: Absolute positioning is selected (1: absolute, 0: relative)
      POS_STW1_Bit09_DirPos : Bool;   // 9: MDI direction selection, positive
      POS_STW1_Bit10_DirNeg : Bool;   // 10: MDI direction selection, negative
      POS_STW1_Bit11_Reserved : Bool;   // 11: Reserved
      POS_STW1_Bit12_Continuous : Bool;   // 12: Continuous transfer (1: continuous setpoint acceptance)
      POS_STW1_Bit13_Reserved : Bool;   // 13: Reserved
      POS_STW1_Bit14_SetupOrPositioning : Bool;   // 14: Toggling the axis operating mode (1: Set up, 0: Positioning)
      POS_STW1_Bit15_ActivateMDI : Bool;   // 15: The converter receives its position setpoint from an
      POS_STW2_Bit00_ActivateFollowUp : Bool;   // 0: Continuously corrects the position setpoint to
      POS_STW2_Bit01_SetRefPoint : Bool;   // 1: Set reference point (0->1: set)
      POS_STW2_Bit02_RefCam : Bool;   // 2: Reference cam active
      POS_STW2_Bit03_AdjustEncoder : Bool;   // 3: Encoder adjustment (0->1: adjust)
      POS_STW2_Bit04_Reserved : Bool;   // 4: Reserved
      POS_STW2_Bit05_JogIncrementalOrVelocity : Bool;   // 5: Jogging mode (1: incremental, 0: velocity)
      POS_STW2_Bit06_Reserved : Bool;   // 6: Reserved
      POS_STW2_Bit07_Reserved : Bool;   // 7: Reserved
      POS_STW2_Bit08_RefType : Bool;   // 8: Referencing type selection (1: flying homing 0: homing approach)
      POS_STW2_Bit09_RefNegDir : Bool;   // 9: Start search for reference direction (1: negative dir, 0: positive dir)
      POS_STW2_Bit10_MeasProbe2 : Bool;   // 10: Measuring probe 2 is activated
      POS_STW2_Bit11_MeasProbeEdge : Bool;   // 11: Falling edge of measuring probe
      POS_STW2_Bit12_Reserved : Bool;   // 12: Reserved
      POS_STW2_Bit13_Reserved : Bool;   // 13: Reserved
      POS_STW2_Bit14_SWLimit : Bool;   // 14: Software limit switch activation
      POS_STW2_Bit15_StopCam : Bool;   // 15: STOP cam active
      STW2_Bit00_Reserved : Bool;   // 0: Reserved
      STW2_Bit01_Reserved : Bool;   // 1: Reserved
      STW2_Bit02_Reserved : Bool;   // 2: Reserved
      STW2_Bit03_Reserved : Bool;   // 3: Reserved
      STW2_Bit04_Reserved : Bool;   // 4: Reserved
      STW2_Bit05_Reserved : Bool;   // 5: Reserved
      STW2_Bit06_Reserved : Bool;   // 6: Reserved
      STW2_Bit07_Reserved : Bool;   // 7: Reserved
      STW2_Bit08_Reserved : Bool;   // 8: Reserved
      STW2_Bit09_Reserved : Bool;   // 9: Reserved
      STW2_Bit10_Reserved : Bool;   // 10: Reserved
      STW2_Bit11_Reserved : Bool;   // 11: Reserved
      STW2_Bit12_Reserved : Bool;   // 12: Reserved
      STW2_Bit13_Reserved : Bool;   // 13: Reserved
      STW2_Bit14_Reserved : Bool;   // 14: Reserved
      STW2_Bit15_Reserved : Bool;   // 15: Reserved
      Override : Int;   // Velocity override [0-4000h = 0-16384 = 0-100%]
      MDI_TARPOS : Real;   // MDI target position
      MDI_VELOCITY : Real;   // MDI velocity
      MDI_ACC : Real;   // MDI acceleration override
      MDI_DEC : Real;   // MDI deceleration override
      Reserved : Real;   // Reserved for future use
      REF_COORDINATE : Real;   // EPOS home position signal
   END_STRUCT;

END_TYPE

TYPE "UDT_S210_HW_Input"
VERSION : 0.1
   STRUCT
      ZSW1_Bit00_ReadyOn : Bool;   // 0: Ready for switching on
      ZSW1_Bit01_Ready : Bool;   // 1: Ready for operation
      ZSW1_Bit02_Enabled : Bool;   // 2: Operation enabled
      ZSW1_Bit03_Fault : Bool;   // 3: Fault present (1: fault)
      ZSW1_Bit04_Off2Inactive : Bool;   // 4: OFF2 inactive (0: active)
      ZSW1_Bit05_Off3Inactive : Bool;   // 5: OFF3 inactive (0: active)
      ZSW1_Bit06_Inhibit : Bool;   // 6: Switching on inhibited
      ZSW1_Bit07_Alarm : Bool;   // 7: Alarm present (1: alarm)
      ZSW1_Bit08_FollowingOK : Bool;   // 8: Following error within tolerance
      ZSW1_Bit09_Control : Bool;   // 9: Control requested
      ZSW1_Bit10_TargetReached : Bool;   // 10: Target position reached
      ZSW1_Bit11_HomeSet : Bool;   // 11: Home position set
      ZSW1_Bit12_AckActive : Bool;   // 12: Acknowledgement traversing block activated
      ZSW1_Bit13_SetpointFixed : Bool;   // 13: Setpoint fixed
      ZSW1_Bit14_AxisAccel : Bool;   // 14: Axis accelerated
      ZSW1_Bit15_AxisDecel : Bool;   // 15: Axis decelerated
      POS_ZSW1_Bit00_Active0 : Bool;   // 0: Active traversing block, bit 0
      POS_ZSW1_Bit01_Active1 : Bool;   // 1: Active traversing block, bit 1
      POS_ZSW1_Bit02_Active2 : Bool;   // 2: Active traversing block, bit 2
      POS_ZSW1_Bit03_Active3 : Bool;   // 3: Active traversing block, bit 3
      POS_ZSW1_Bit04_Active4 : Bool;   // 4: Active traversing block, bit 4
      POS_ZSW1_Bit05_Active5 : Bool;   // 5: Active traversing block, bit 5
      POS_ZSW1_Bit06_Reserved : Bool;   // 6: Reserved
      POS_ZSW1_Bit07_ReleaseBrake : Bool;   // 7: The converter opens the holding brake
      POS_ZSW1_Bit08_StopCamMinus : Bool;   // 8: STOP cam minus active
      POS_ZSW1_Bit09_StopCamPlus : Bool;   // 9: STOP cam plus active
      POS_ZSW1_Bit10_JogActive : Bool;   // 10: Jogging active (r2669.0)
      POS_ZSW1_Bit11_RefApproach : Bool;   // 11: Reference point approach active (r2669.1)
      POS_ZSW1_Bit12_FlyingHoming : Bool;   // 12: Homes when passing the reference cam
      POS_ZSW1_Bit13_Traversing : Bool;   // 13: Traversing block active (r2669.2)
      POS_ZSW1_Bit14_Setup : Bool;   // 14: Setup active (r2669.4)
      POS_ZSW1_Bit15_MDI : Bool;   // 15: MDI active
      POS_ZSW2_Bit00_Tracking : Bool;   // 0: Tracking mode active
      POS_ZSW2_Bit01_VelLimit : Bool;   // 1: Velocity limiting active
      POS_ZSW2_Bit02_TargetReached : Bool;   // 2: Target position reached (r2683.3)
      POS_ZSW2_Bit03_PrintMark : Bool;   // 3: Printing mark outside outer window
      POS_ZSW2_Bit04_Forward : Bool;   // 4: Axis moves forward
      POS_ZSW2_Bit05_Backward : Bool;   // 5: Axis moves backward
      POS_ZSW2_Bit06_SWLimitMinus : Bool;   // 6: Software limit switch minus reached
      POS_ZSW2_Bit07_SWLimitPlus : Bool;   // 7: Software limit switch plus reached
      POS_ZSW2_Bit08_Cam1 : Bool;   // 8: Position actual value <= cam switching position 1
      POS_ZSW2_Bit09_Cam2 : Bool;   // 9: Position actual value <= cam switching position 2
      POS_ZSW2_Bit10_Output1 : Bool;   // 10: Direct output 1 via traversing block
      POS_ZSW2_Bit11_Output2 : Bool;   // 11: Direct output 2 via traversing block
      POS_ZSW2_Bit12_FixedStop : Bool;   // 12: Fixed stop reached
      POS_ZSW2_Bit13_Clamping : Bool;   // 13: Fixed stop clamping torque reached
      POS_ZSW2_Bit14_TravelFixed : Bool;   // 14: Travel to fixed stop active
      POS_ZSW2_Bit15_TraversingCmd : Bool;   // 15: Traversing command active
      ZSW2_Bit00_Reserved : Bool;   // 0: Reserved
      ZSW2_Bit01_Reserved : Bool;   // 1: Reserved
      ZSW2_Bit02_Reserved : Bool;   // 2: Reserved
      ZSW2_Bit03_Reserved : Bool;   // 3: Reserved
      ZSW2_Bit04_Reserved : Bool;   // 4: Reserved
      ZSW2_Bit05_Reserved : Bool;   // 5: Reserved
      ZSW2_Bit06_Reserved : Bool;   // 6: Reserved
      ZSW2_Bit07_Reserved : Bool;   // 7: Reserved
      ZSW2_Bit08_Reserved : Bool;   // 8: Reserved
      ZSW2_Bit09_Reserved : Bool;   // 9: Reserved
      ZSW2_Bit10_Reserved : Bool;   // 10: Reserved
      ZSW2_Bit11_Reserved : Bool;   // 11: Reserved
      ZSW2_Bit12_Reserved : Bool;   // 12: Reserved
      ZSW2_Bit13_Reserved : Bool;   // 13: Reserved
      ZSW2_Bit14_Reserved : Bool;   // 14: Reserved
      ZSW2_Bit15_Reserved : Bool;   // 15: Reserved
      Reserved : Int;   // Reserved
      XIST : Real;   // Position actual value
      VIST : Real;   // Velocity actual value
      MELDW_Bit00_PositioningAbsolute : Bool;   // 0: Positioning mode (1: absolute, 0: relative)
      MELDW_Bit01_AbsolutePositiveDir : Bool;   // 1: Absolute positioning for rotary axis in the positive direction
      MELDW_Bit02_AbsoluteNegativeDir : Bool;   // 2: Absolute positioning for rotary axes in negative direction
      MELDW_Bit03_Reserved : Bool;   // 3: Reserved
      MELDW_Bit04_Reserved : Bool;   // 4: Reserved
      MELDW_Bit05_Reserved : Bool;   // 5: Reserved
      MELDW_Bit06_Reserved : Bool;   // 6: Reserved
      MELDW_Bit07_Reserved : Bool;   // 7: Reserved
      MELDW_Bit08_Reserved : Bool;   // 8: Reserved
      MELDW_Bit09_Reserved : Bool;   // 9: Reserved
      MELDW_Bit10_Reserved : Bool;   // 10: Reserved
      MELDW_Bit11_Reserved : Bool;   // 11: Reserved
      MELDW_Bit12_Reserved : Bool;   // 12: Reserved
      MELDW_Bit13_Reserved : Bool;   // 13: Reserved
      MELDW_Bit14_Reserved : Bool;   // 14: Reserved
      MELDW_Bit15_Reserved : Bool;   // 15: Reserved
      FaultCode : Word;   // Fault code (0: no fault)
      AlarmCode : Word;   // Alarm code (0: no alarm)
      ZSW_S210_Bit00_DI0 : Bool;   // 0: Digital input 0 status
      ZSW_S210_Bit01_DI1 : Bool;   // 1: Digital input 1 status
      ZSW_S210_Bit02_DI2 : Bool;   // 2: Digital input 2 status
      ZSW_S210_Bit03_DI3 : Bool;   // 3: Digital input 3 status
      ZSW_S210_Bit04_DI4 : Bool;   // 4: Digital input 4 status
      ZSW_S210_Bit05_Reserved : Bool;   // 5: Reserved
      ZSW_S210_Bit06_Reserved : Bool;   // 6: Reserved
      ZSW_S210_Bit07_Reserved : Bool;   // 7: Reserved
      ZSW_S210_Bit08_Reserved : Bool;   // 8: Reserved
      ZSW_S210_Bit09_Reserved : Bool;   // 9: Reserved
      ZSW_S210_Bit10_Reserved : Bool;   // 10: Reserved
      ZSW_S210_Bit11_Reserved : Bool;   // 11: Reserved
      ZSW_S210_Bit12_Reserved : Bool;   // 12: Reserved
      ZSW_S210_Bit13_Reserved : Bool;   // 13: Reserved
      ZSW_S210_Bit14_Reserved : Bool;   // 14: Reserved
      ZSW_S210_Bit15_Reserved : Bool;   // 15: Reserved
      DCLinkVoltage : Int;   // DC link voltage [V]
      ActualCurrent : Int;   // Actual current [0.1A]
      ActivePower : Int;   // Active power [W]
      TorqueUtilization : Int;   // Torque utilization [%]
      MotorUtilization : Int;   // Motor utilization thermal [%]
   END_STRUCT;

END_TYPE

TYPE "UDT_Commen_Setting"
TITLE = UDT_Commen_Setting
VERSION : 0.1
//# Block Info
//- Title:            UDT_Commen_Setting
//- Comment/Function: ---
//- Library/Family:   APS
//- Author:           Jay Liu
//- Tested with:      ---
//- Engineering:      TIA Portal V20
//- Restrictions:     ---
//- Requirements:     ---
//
//# History
// |Version  | Date       | Author                 | Description                   |
// |---------|------------|------------------------|------------------------------ |
// |01.00.00 | 2026-01-22 | Jay Liu                | First released version        |
   STRUCT
      Auto_Start : Bool;
      Alarms_Need_ACK : Bool;
      Disable_Energy_Saving : Bool;
      PECTrigger_During_E_Save : Bool;
      Disable_PEC_Blockage : Bool;
      Log_Level : Int;
      Max_Product_Length : Int;   // [cm]
   END_STRUCT;

END_TYPE

TYPE "UDT_Conv_S210_Diagnostics"
VERSION : 0.1
   STRUCT
      RTS : Bool;   // Section ready to send item
      TIP : Bool;   // Section transfer in porgress
      Downstream_RTR : Bool;   // Downstream section ready to receive item
      Items_Count : UDInt;   // Count of items passed
      Displacement : Int;   // [mm/scan] Conveyor movement distance
      Hardware { S7_SetPoint := 'False'} : "UDT_S210_HW_Diagnostics";
   END_STRUCT;

END_TYPE

TYPE "UDT_Conv_S210_Setting"
VERSION : 0.1
   STRUCT
      PE1 { S7_SetPoint := 'False'} : "UDT_PEC_Position_Setting";
      PE2 : "UDT_PEC_Trigger_Setting";
      Flow_Control : "UDT_Flow_Control_Setting";
      Base_Conveyor : "UDT_Base_Conveyor_Setting";
      Hardware : "UDT_S210_Speed_Setting" := (1200, (), (), (), (), (), (), (), (), (), (), ());
   END_STRUCT;

END_TYPE

TYPE "UDT_NBS_Setting"
VERSION : 0.1
   STRUCT
      StartUp_Delay : Int;   // [ms]
      Dieback_Delay : Int;   // [ms]
   END_STRUCT;

END_TYPE

TYPE "UDT_ADTA_Setting"
VERSION : 0.1
   STRUCT
      StartUp_Delay : Int;   // [ms]
      Dieback_Delay : Int;   // [ms]
   END_STRUCT;

END_TYPE

TYPE "UDT_RLS_Setting"
VERSION : 0.1
   STRUCT
      StartUp_Delay : Int;   // [ms]
      Dieback_Delay : Int;   // [ms]
   END_STRUCT;

END_TYPE

TYPE "UDT_Conv_G115D_Setting"
VERSION : 0.1
   STRUCT
      PE1 { S7_SetPoint := 'False'} : "UDT_PEC_Position_Setting";
      PE2 : "UDT_PEC_Trigger_Setting";
      Flow_Control : "UDT_Flow_Control_Setting";
      Base_Conveyor : "UDT_Base_Conveyor_Setting";
      Hardware : "UDT_G115D_Setting" := (1200, (), (), (), 4000, 4000, 2000, 10000, (), (), ());
   END_STRUCT;

END_TYPE

TYPE "UDT_IOLink_Master_Setting"
VERSION : 0.1
   STRUCT
      Bypass_Time : Int;   // [ms]
   END_STRUCT;

END_TYPE

TYPE "UDT_Accmulation_Setting"
VERSION : 0.1
   STRUCT
      Gap : DInt;   // [mm]
      Cleanup_Distance : DInt;   // [mm]
      Waiting_Timeout : DInt;   // [s]
      Max_Count : Int;
   END_STRUCT;

END_TYPE

TYPE "UDT_Conv_Triple_G115D_Setting"
VERSION : 0.1
   STRUCT
      PE1 { S7_SetPoint := 'False'} : "UDT_PEC_Position_Setting";
      PE2 : "UDT_PEC_Trigger_Setting";
      Flow_Control : "UDT_Flow_Control_Setting";
      Base_Conveyor : "UDT_Base_Conveyor_Setting";
      Hardware_U01 : "UDT_G115D_Setting" := (1000, (), (), (), 4000, 4000, 2000, 10000, (), (), ());
      Hardware_U02 : "UDT_G115D_Setting";
      Hardware_U03 : "UDT_G115D_Setting";
   END_STRUCT;

END_TYPE

TYPE "UDT_Merge_3_To_1_Setting"
VERSION : 0.1
   STRUCT
      Line1_Infeed_Delay : Int;
      Line1_Waiting_Delay : Int;
      Line2_Infeed_Delay : Int;
      Line2_Waiting_Delay : Int;
      Line3_Infeed_Delay : Int;
      Line3_Waiting_Delay : Int;
   END_STRUCT;

END_TYPE

TYPE "UDT_MultiControl_HW_Output"
VERSION : 0.1
   STRUCT
      Output1 : Bool;
      Output2 : Bool;
      Output3 : Bool;
      Output4 : Bool;
      MotorSpeed_RD1 : SInt;
      MotorSpeed_RD2 : SInt;
      MotorSpeed_RD3 : SInt;
      MotorSpeed_RD4 : SInt;
   END_STRUCT;

END_TYPE

TYPE "UDT_Conv_Dual_G115D_Setting"
VERSION : 0.1
   STRUCT
      PE1 { S7_SetPoint := 'False'} : "UDT_PEC_Position_Setting";
      PE2 : "UDT_PEC_Trigger_Setting";
      Flow_Control : "UDT_Flow_Control_Setting";
      Base_Conveyor : "UDT_Base_Conveyor_Setting";
      Hardware_U01 : "UDT_G115D_Setting" := (1000, (), (), (), 4000, 4000, 2000, 10000, (), (), ());
      Hardware_U02 : "UDT_G115D_Setting";
   END_STRUCT;

END_TYPE

TYPE "UDT_Induct_On_Gap_Setting"
VERSION : 0.1
   STRUCT
      Induct_Position : DInt;
      Gap_Length : Int;
      Max_Item_Length : Int;
   END_STRUCT;

END_TYPE

TYPE "UDT_Conv_Multiple_S210_Setting"
VERSION : 0.1
   STRUCT
      PE1 { S7_SetPoint := 'False'} : "UDT_PEC_Position_Setting";
      PE2 : "UDT_PEC_Trigger_Setting";
      Flow_Control : "UDT_Flow_Control_Setting";
      Base_Conveyor : "UDT_Base_Conveyor_Setting";
      Hardware_U01 : "UDT_S210_Speed_Setting";
      Hardware_U02 : "UDT_S210_Speed_Setting";
      Hardware_U03 : "UDT_S210_Speed_Setting";
      Hardware_U04 : "UDT_S210_Speed_Setting";
      Hardware_U05 : "UDT_S210_Speed_Setting";
      Hardware_U06 : "UDT_S210_Speed_Setting";
      Hardware_U07 : "UDT_S210_Speed_Setting";
      Hardware_U08 : "UDT_S210_Speed_Setting";
      Hardware_U09 : "UDT_S210_Speed_Setting";
      Hardware_U10 : "UDT_S210_Speed_Setting";
   END_STRUCT;

END_TYPE

TYPE "UDT_Merge_2_To_1_Setting"
VERSION : 0.1
   STRUCT
      Line1_Infeed_Delay : Int;
      Line1_Waiting_Delay : Int;
      Line2_Infeed_Delay : Int;
      Line2_Waiting_Delay : Int;
   END_STRUCT;

END_TYPE

TYPE "UDT_Conv_MultiControl_Setting"
VERSION : 0.1
   STRUCT
      PE1 { S7_SetPoint := 'False'} : "UDT_PEC_Position_Setting";
      PE2 : "UDT_PEC_Trigger_Setting";
      Flow_Control : "UDT_Flow_Control_Setting";
      Base_Conveyor : "UDT_Base_Conveyor_Setting";
      Hardware_U01 : "UDT_MultiControl_Setting";
      Hardware_U02 : "UDT_MultiControl_Setting";
      Hardware_U03 : "UDT_MultiControl_Setting";
      Hardware_U04 : "UDT_MultiControl_Setting";
   END_STRUCT;

END_TYPE

TYPE "UDT_Conv_SWS_Setting"
VERSION : 0.1
   STRUCT
      Decision : "UDT_Divert_Decision_Setting";
      Divert : "UDT_SWS_Divert_Setting" := ((), 1, 1, 300, (), (), (), 170, 170, 170, 170, 170);
      Base_Conveyor : "UDT_Base_Conveyor_Setting";
      Roller_Interface : "UDT_SWS_Roller_Interface_Setting";
      Hardware : "UDT_SWS_Hardware_Setting";
   END_STRUCT;

END_TYPE

TYPE "UDT_Chute_Setting"
VERSION : 0.1
   STRUCT
      PEC_Full { S7_SetPoint := 'False'} : "UDT_PEC_Trigger_Setting" := (3000, 50, 50, TRUE, (), FALSE);
   END_STRUCT;

END_TYPE

TYPE "UDT_Track_Setting"
VERSION : 0.1
   STRUCT
      Measure_Length : Bool;
      Update_Position : DInt;
      Open_Window : DInt := 200;
      Close_Window : DInt := 200;
      Package_Range : Int;
      Num_MIssing_Error : Int := 5;
      Upd_Perf_WN_Level : Int := 80;
      Localtion : String[10];
   END_STRUCT;

END_TYPE

TYPE "UDT_MultiControl_HW_Interface"
VERSION : 0.1
   STRUCT
      Input { S7_SetPoint := 'False'} : "UDT_MultiControl_HW_Input";
      Output { S7_SetPoint := 'False'} : "UDT_MultiControl_HW_Output";
   END_STRUCT;

END_TYPE

TYPE "UDT_SWS_Roller_Module_Status"
VERSION : 0.1
   STRUCT
      WN_Modbus_Com_Error : Bool;
      WN_Motor_NotConnected : Bool;
      WN_Motor_Blockage : Bool;
      WN_Motor_NotHealthy : Bool;
      Spare_0_4 : Bool;
      Spare_0_5 : Bool;
      Spare_0_6 : Bool;
      Spare_0_7 : Bool;
      Spare_1_0 : Bool;
      Spare_1_1 : Bool;
      Spare_1_2 : Bool;
      Spare_1_3 : Bool;
      Spare_1_4 : Bool;
      Spare_1_5 : Bool;
      Spare_1_6 : Bool;
      Spare_1_7 : Bool;
   END_STRUCT;

END_TYPE

TYPE "UDT_SWS_Roller_IO"
VERSION : 0.1
   STRUCT
      Input : Struct
         Alarm : Bool;
      END_STRUCT;
      Output : Struct
         Direction : Bool;
         Array1_Speed1 : Bool;
         Array1_Speed2 : Bool;
         Array2_Speed1 : Bool;
         Array2_Speed2 : Bool;
         Array3_Speed1 : Bool;
         Array3_Speed2 : Bool;
         Array4_Speed1 : Bool;
         Array4_Speed2 : Bool;
         Array5_Speed1 : Bool;
         Array5_Speed2 : Bool;
         Array6_Speed1 : Bool;
         Array6_Speed2 : Bool;
         Array7_Speed1 : Bool;
         Array7_Speed2 : Bool;
         Array8_Speed1 : Bool;
         Array8_Speed2 : Bool;
         Array9_Speed1 : Bool;
         Array9_Speed2 : Bool;
      END_STRUCT;
   END_STRUCT;

END_TYPE

TYPE "UDT_SWS_Servo_Command"
VERSION : 0.1
   STRUCT
      Man_Disable_Axis : Bool;   // Maintenance - Disable axis enable
      Man_Home : Bool;   // Maintenance - Adujst encoder
      Man_Jog_Left : Bool;   // Maintenance - Jog to divert left
      Man_Jog_Right : Bool;   // Maintenance - Jog to divert right
      Man_Save_Parameter : Bool;
   END_STRUCT;

END_TYPE

FUNCTION "FC_Delay_On_Accumulator" : Void
{ S7_Optimized_Access := 'TRUE' }
VERSION : 0.1
   VAR_INPUT
      i_CMD_Start : Bool;
      i_Enable_Dly : Bool;
      i_CFG_Target : Int;
      i_Cycle_Count : Int;
   END_VAR

   VAR_OUTPUT
      o_Delay_Finish : Bool;
   END_VAR

   VAR_IN_OUT
      io_Setpoint : Int;
   END_VAR


BEGIN
	// Init time value
	IF NOT #i_CMD_Start THEN
	    #io_Setpoint := 0;
	END_IF;

	// Detect result
	#o_Delay_Finish := #i_CMD_Start AND #io_Setpoint >= #i_CFG_Target;

	// Count time value
	IF #i_CMD_Start THEN
	    IF #i_Enable_Dly THEN
	        #io_Setpoint := #io_Setpoint + #i_Cycle_Count;
	    END_IF;
	    IF #io_Setpoint > #i_CFG_Target THEN
	        #io_Setpoint := #i_CFG_Target;
	    END_IF;
	END_IF;
END_FUNCTION

TYPE "UDT_NT100_Output"
VERSION : 0.1
   STRUCT
      APP_HS_TX_CMD : Bool;
      APP_HS_RX_ACK : Bool;
      Spare_0_2 : Bool;
      Spare_0_3 : Bool;
      Spare_0_4 : Bool;
      Spare_0_5 : Bool;
      APP_HS_TX_ENABLE_CMD : Bool;
      APP_HS_RX_ENABLE_CMD : Bool;
      Spare_1_0 : Bool;
      Spare_1_1 : Bool;
      Spare_1_2 : Bool;
      Spare_1_3 : Bool;
      Spare_1_4 : Bool;
      Spare_1_5 : Bool;
      Spare_1_6 : Bool;
      APP_HS_RESET_CMD : Bool;
      Spare_Word_1 : Word;
      User_Data_Length : UDInt;
      User_Data : Array[1..56] of Byte;
   END_STRUCT;

END_TYPE

FUNCTION_BLOCK "FB_SINA_Save_Parameter"
{ S7_Optimized_Access := 'TRUE' }
VERSION : 0.1
   VAR_INPUT
      i_Trigger : Bool;
      i_VFD_Type : Int;   // 1: G115D 2: S210
      i_HW_ID : HW_ANY;
   END_VAR

   VAR_OUTPUT
      o_Ready : Bool;
      o_Busy : Bool;
      o_Done : Bool;
      o_Error : Bool;
   END_VAR

   VAR
      s_SinaParaS {InstructionName := 'SinaParaS'; LibVersion := '1.1'} : SinaParaS;
      s_Copy_Trigger { S7_SetPoint := 'True'} : Bool;
      s_Excute : Bool;
   END_VAR

   VAR_TEMP
      t_Parameter : UInt;
   END_VAR

   VAR CONSTANT
      C_G115D_P_INDEX : UInt := 971;
      C_S210_P_INDEX : UInt := 977;
   END_VAR


BEGIN
	IF #i_VFD_Type = 1 THEN
	    #t_Parameter := #C_G115D_P_INDEX;
	ELSIF #i_VFD_Type = 2 THEN
	    #t_Parameter := #C_S210_P_INDEX;
	ELSE
	    RETURN;
	END_IF;

	IF #i_Trigger AND NOT #s_Copy_Trigger THEN
	    #s_Excute := TRUE;
	END_IF;

	#s_SinaParaS(Start       := #s_Excute,
	             ReadWrite   := TRUE,
	             Parameter   := #t_Parameter,
	             Index       := 0,
	             ValueWrite1 := 1.0,
	             AxisNo      := 1,
	             hardwareId  := #i_HW_ID,
	             Ready       => #o_Ready,
	             Busy        => #o_Busy,
	             Done        => #o_Done,
	             Error       => #o_Error);

	IF NOT #o_Busy THEN
	    #s_Excute := FALSE;
	END_IF;

	#s_Copy_Trigger := #i_Trigger;
END_FUNCTION_BLOCK

FUNCTION "FC_SWS_Convert_Motor_Status" : Void
{ S7_Optimized_Access := 'TRUE' }
VERSION : 0.1
   VAR_INPUT
      i_Status_Byte_1 : Byte;
      i_Status_Byte_2 : Byte;
   END_VAR

   VAR_OUTPUT
      o_Motor_Status : "UDT_SWS_Roller_Module_Motor_Status";
   END_VAR

   VAR_TEMP
      t_Status_Word : Word;
   END_VAR


BEGIN
	#t_Status_Word.%B0 := #i_Status_Byte_1;
	#t_Status_Word.%B1 := #i_Status_Byte_2;

	IF #t_Status_Word = 16#FFFF THEN
	    #o_Motor_Status.None := TRUE;
	    #o_Motor_Status.NotConnected := FALSE;
	    #o_Motor_Status.Blockage := FALSE;
	    #o_Motor_Status.OK := FALSE;
	ELSIF #t_Status_Word = 16#80C0 THEN
	    #o_Motor_Status.None := FALSE;
	    #o_Motor_Status.NotConnected := TRUE;
	    #o_Motor_Status.Blockage := FALSE;
	    #o_Motor_Status.OK := FALSE;
	ELSIF #t_Status_Word = 16#0040 THEN
	    #o_Motor_Status.None := FALSE;
	    #o_Motor_Status.NotConnected := FALSE;
	    #o_Motor_Status.Blockage := TRUE;
	    #o_Motor_Status.OK := FALSE;
	ELSE
	    #o_Motor_Status.None := FALSE;
	    #o_Motor_Status.NotConnected := FALSE;
	    #o_Motor_Status.Blockage := FALSE;
	    #o_Motor_Status.OK := TRUE;
	END_IF;

END_FUNCTION

TYPE "UDT_NT100_Input"
VERSION : 0.1
   STRUCT
      PROT_HS_TX_ACK : Bool;
      PROT_HS_RX_CMD : Bool;
      Spare_0_2 : Bool;
      PROT_HS_RUN_IND : Bool;
      PROT_HS_TX_ERROR_IND : Bool;
      PROT_HS_RX_ERROR_IND : Bool;
      PROT_HS_TX_ENABLE_ACK : Bool;
      PROT_HS_RX_ENABLE_ACK : Bool;
      Spare_1_0 : Bool;
      Spare_1_1 : Bool;
      Spare_1_2 : Bool;
      Spare_1_3 : Bool;
      Spare_1_4 : Bool;
      Spare_1_5 : Bool;
      Spare_1_6 : Bool;
      PROT_HS_RESET_ACK : Bool;
      Spare_Word_1 : Word;
      Input_Data_Length : UDInt;
      Recv_Error_Code : DWord;
      Send_Error_Code : DWord;
      Input_Data : Array[1..112] of Byte;
   END_STRUCT;

END_TYPE

TYPE "UDT_SWS_Servo_Status"
VERSION : 0.1
   STRUCT
      ER_PN_NotPresent : Bool;
      ER_PN_Error : Bool;
      OL_Maintenance_Mode : Bool;
      ST_Axis_Enabled : Bool;
      ST_Axis_Position_Reached : Bool;
      ER_Home_Position_Missed : Bool;
      WN_Servo_Warn : Bool;
      ER_Servo_Fault : Bool;
      ER_STO_Active : Bool;
      Spare_1_1 : Bool;
      Spare_1_2 : Bool;
      Spare_1_3 : Bool;
      Spare_1_4 : Bool;
      Spare_1_5 : Bool;
      Spare_1_6 : Bool;
      Spare_1_7 : Bool;
      ST_Act_Position : Real;
      AlarmCode : Word;
      ErrorCode : Word;
   END_STRUCT;

END_TYPE

TYPE "UDT_Flow_Interface"
TITLE = UDT_Flow_Interface
VERSION : 0.1
//Flow interface of each section and unit
//# Block Info
//- Title:            UDT_Flow_Interface
//- Comment/Function: Flow interface of each section and unit
//- Library/Family:   APS
//- Author:           Jay Liu
//- Tested with:      ---
//- Engineering:      TIA Portal V20
//- Restrictions:     ---
//- Requirements:     ---
//
//# History
// |Version  | Date       | Author                 | Description                   |
// |---------|------------|------------------------|------------------------------ |
// |01.00.00 | 2026-01-22 | Jay Liu                | First released version        |
   STRUCT
      Item_at_Handover : Bool;   // [Up -> Down] Item at Handover position
      RTS : Bool;   // [Up -> Down] Ready To Send
      RTR : Bool;   // [Down -> Up] Ready To Receive
      TIP : Bool;   // [Up -> Down] Transfer in progress
      Handover : Bool;   // [Up -> Down] Handover Item
      Operational : Bool;   // [Down -> Up] Section is operational on
      Available : Bool;   // [Down -> Up] Section is available
      Cascade_Startup : Bool;   // [Down -> Up] Cascade start up upstream
      Cascade_Shutdown : Bool;   // [Up -> Down] Cascade shutdown downstream
      Motor_Run : Bool;   // [Down -> Up] Motor is running
      Motor_Stopped : Bool;   // [Down -> Up] Motor is stopped
      Receive_Item : Bool;   // [Down -> Up] Waiting item to the End PEC
      Items : Bool;   // [Down -> Up] Section have items
      PECPosition_Latch : Bool;   // [Up -> Down] PEC Latch at the end
      PECTrigger_Latch : Bool;   // [Up -> Down] PEC Latch on the conveyor
      Data_Sync : Bool;   // [Up -> Down] (One-shot) Hand-Over of data
      Req_Up_Disable_Send : Bool;   // [Down -> Up] Request Disable send new products
      Req_Upstream_Halt : Bool;   // [Down -> Up] Request Halt Upstream
      Req_Down_Reset_E_Saving : Bool;   // [Up -> Down] Request Reset energy saving
      Req_Down_Disable_Receive : Bool;   // [Up -> Down] Request Disable receiving new products
      Req_Downstream_Halt : Bool;   // [Up -> Down] Request Halt Downstream
      Speed : Int;   // [mm/s] Speed setpoint
      Displacement : Int;   // [mm] Cycle displacement
      Data : Int;   // Tracking Data
   END_STRUCT;

END_TYPE

DATA_BLOCK "DB_Diagnostics"
{ S7_Optimized_Access := 'TRUE' }
VERSION : 0.1
NON_RETAIN
   VAR
      Rack : "UDT_IODevice_Diag";
      PNIO_System_100 : "UDT_PNIO_System_Diag";
      GC03_CT01 { S7_SetPoint := 'False'} : "UDT_Scanner_Statistics";
      GC04_CT01 { S7_SetPoint := 'False'} : "UDT_Scanner_Statistics";
      Inbound1_Infeed : "UDT_Mesasuring_Point_Statistics";
      Inbound1_OV : "UDT_Mesasuring_Point_Statistics";
      Inbound1_NonOV : "UDT_Mesasuring_Point_Statistics";
      Inound3_NonOV : "UDT_Mesasuring_Point_Statistics";
      InoundNonOV : "UDT_Mesasuring_Point_Statistics";
      InboundOV_MergeOV : "UDT_Mesasuring_Point_Statistics";
      GC01_FB01 : "UDT_Conv_G115D_Diagnostics";
      GC01_FB02 : "UDT_Conv_G115D_Diagnostics";
      GC01_FB03_Track : "UDT_Track_Statistics";
      GC01_FB03 : "UDT_Conv_G115D_Diagnostics";
      GC01_FB04_Track : "UDT_Track_Statistics";
      GC01_FB04 : "UDT_Conv_S210_Diagnostics";
      GC01_FB05_Track : "UDT_Track_Statistics";
      GC01_FB05 : "UDT_Conv_S210_Diagnostics";
      DT01 : "UDT_Divert_Statistics";
      GC01_RC06_Track : "UDT_Track_Statistics";
      GC01_RC06 : "UDT_Conv_MultiControl_Diagnostics";
      GC01_FB07 : "UDT_Conv_G115D_Diagnostics";
      GC01_FB08 : "UDT_Conv_G115D_Diagnostics";
      GC01_RC09 : "UDT_Conv_MultiControl_Diagnostics";
      GC01_RC09_Track : "UDT_Track_Statistics";
      GC01_RC10 : "UDT_Conv_MultiControl_Diagnostics";
      GC01_RC40 : "UDT_Conv_MultiControl_Diagnostics";
      GC01_SK11 : "UDT_Conv_G115D_Diagnostics";
      GC01_FB12 : "UDT_Conv_S210_Diagnostics";
      GC01_FB13 : "UDT_Conv_S210_Diagnostics";
      GC01_FB14 : "UDT_Conv_S210_Diagnostics";
      GC01_FB15 : "UDT_Conv_G115D_Diagnostics";
      GC01_FB16 : "UDT_Conv_G115D_Diagnostics";
      GC01_FB17 : "UDT_Conv_G115D_Diagnostics";
      GC01_FB18 : "UDT_Conv_G115D_Diagnostics";
      GC01_FB19 : "UDT_Conv_G115D_Diagnostics";
      GC01_FB20 : "UDT_Conv_G115D_Diagnostics";
      GC01_FB21 : "UDT_Conv_G115D_Diagnostics";
      GC01_FB22 : "UDT_Conv_G115D_Diagnostics";
      GC01_FB23 : "UDT_Conv_G115D_Diagnostics";
      GC01_FB24 : "UDT_Conv_G115D_Diagnostics";
      GC01_FB25 : "UDT_Conv_G115D_Diagnostics";
      GC01_FB26 : "UDT_Conv_G115D_Diagnostics";
      GC01_FB27 : "UDT_Conv_G115D_Diagnostics";
      GC01_FB28 : "UDT_Conv_S210_Diagnostics";
      GC01_FB29 : "UDT_Conv_S210_Diagnostics";
      GC01_FB30 : "UDT_Conv_S210_Diagnostics";
      GC01_FB31 : "UDT_Conv_S210_Diagnostics";
      GC01_FB32 : "UDT_Conv_G115D_Diagnostics";
      GC02_FB01 : "UDT_Conv_G115D_Diagnostics";
      GC02_FB02 : "UDT_Conv_G115D_Diagnostics";
      GC02_FB03_Track : "UDT_Track_Statistics";
      GC02_FB03 : "UDT_Conv_S210_Diagnostics";
      GC02_FB04_Track : "UDT_Track_Statistics";
      GC02_FB04 : "UDT_Conv_S210_Diagnostics";
      DT02 : "UDT_Divert_Statistics";
      GC02_RC05_Track : "UDT_Track_Statistics";
      GC02_RC05 : "UDT_Conv_MultiControl_Diagnostics";
      GC02_FB06 : "UDT_Conv_G115D_Diagnostics";
      GC02_FB07 : "UDT_Conv_G115D_Diagnostics";
      GC02_FB08_Track : "UDT_Track_Statistics";
      GC02_FB08 : "UDT_Conv_G115D_Diagnostics";
      GC02_FB09 : "UDT_Conv_G115D_Diagnostics";
      GC02_FB10 : "UDT_Conv_G115D_Diagnostics";
      GC02_FB11 : "UDT_Conv_G115D_Diagnostics";
      GC02_FB12 : "UDT_Conv_G115D_Diagnostics";
      GC02_FB13 : "UDT_Conv_G115D_Diagnostics";
      GC02_FB14 : "UDT_Conv_G115D_Diagnostics";
      GC02_SK15 : "UDT_Conv_G115D_Diagnostics";
      GC02_FB16 : "UDT_Conv_S210_Diagnostics";
      GC02_FB17 : "UDT_Conv_S210_Diagnostics";
      GC02_FB18 : "UDT_Conv_S210_Diagnostics";
      GC03_RC01 : "UDT_Conv_MultiControl_Diagnostics";
      GC03_RC40 : "UDT_Conv_MultiControl_Diagnostics";
      GC03_RC02 : "UDT_Conv_MultiControl_Diagnostics";
      GC03_RC03 : "UDT_Conv_MultiControl_Diagnostics";
      GC03_RC41 : "UDT_Conv_MultiControl_Diagnostics";
      GC03_RC04 : "UDT_Conv_MultiControl_Diagnostics";
      GC03_HB05 : "UDT_Conv_Multiple_S210_Diagnostics";
      GC03_FB06 : "UDT_Conv_G115D_Diagnostics";
      GC03_FB42 : "UDT_Conv_G115D_Diagnostics";
      GC03_FB07 : "UDT_Conv_G115D_Diagnostics";
      GC03_FB08_Track : "UDT_Track_Statistics";
      GC03_FB08 : "UDT_Conv_G115D_Diagnostics";
      GC03_FB09_Track : "UDT_Track_Statistics";
      GC03_FB09 : "UDT_Conv_G115D_Diagnostics";
      GC03_FB10 : "UDT_Conv_S210_Diagnostics";
      GC03_FB11_Track : "UDT_Track_Statistics";
      GC03_FB11 : "UDT_Conv_S210_Diagnostics";
      DT03 : "UDT_Divert_Statistics";
      GC03_CH01 : "UDT_Chute_Statistics";
      GC03_RC12_Track : "UDT_Track_Statistics";
      GC03_RC12 : "UDT_Conv_MultiControl_Diagnostics";
      GC03_FB13 : "UDT_Conv_G115D_Diagnostics";
      GC03_FB14 : "UDT_Conv_S210_Diagnostics";
      GC03_FB15 : "UDT_Conv_S210_Diagnostics";
      GC03_FB16 : "UDT_Conv_S210_Diagnostics";
      GC03_FB17 : "UDT_Conv_S210_Diagnostics";
      GC03_FB18 : "UDT_Conv_G115D_Diagnostics";
      GC03_RC19 : "UDT_Conv_G115D_Diagnostics";
      GC03_RC20 : "UDT_Conv_MultiControl_Diagnostics";
      GC03_FB21 : "UDT_Conv_G115D_Diagnostics";
      GC03_FB22 : "UDT_Conv_G115D_Diagnostics";
      GC03_FB23 : "UDT_Conv_G115D_Diagnostics";
      GC03_FB24 : "UDT_Conv_G115D_Diagnostics";
      GC03_FB25 : "UDT_Conv_G115D_Diagnostics";
      GC03_FB26 : "UDT_Conv_G115D_Diagnostics";
      GC03_FB27 : "UDT_Conv_G115D_Diagnostics";
      GC03_FB28 : "UDT_Conv_G115D_Diagnostics";
      GC03_FB29 : "UDT_Conv_G115D_Diagnostics";
      GC03_FB30 : "UDT_Conv_G115D_Diagnostics";
      GC03_FB31 : "UDT_Conv_G115D_Diagnostics";
      GC03_FB32 : "UDT_Conv_G115D_Diagnostics";
      GC03_RC33_Track : "UDT_Track_Statistics";
      GC03_RC33 : "UDT_Conv_Dual_G115D_Diagnostics";
      GC04_FB04 : "UDT_Conv_G115D_Diagnostics";
      GC04_FB05 : "UDT_Conv_G115D_Diagnostics";
      GC04_FB06 : "UDT_Conv_G115D_Diagnostics";
      GC04_FB07 : "UDT_Conv_G115D_Diagnostics";
      GC04_FB08 : "UDT_Conv_G115D_Diagnostics";
      GC04_FB09_Track : "UDT_Track_Statistics";
      GC04_FB09 : "UDT_Conv_G115D_Diagnostics";
      GC04_FB10 : "UDT_Conv_S210_Diagnostics";
      GC04_FB11_Track : "UDT_Track_Statistics";
      GC04_FB11 : "UDT_Conv_S210_Diagnostics";
      DT04 : "UDT_Divert_Statistics";
      GC04_CH01 : "UDT_Chute_Statistics";
      GC04_FB12 : "UDT_Conv_G115D_Diagnostics";
      GC04_FB13_Track : "UDT_Track_Statistics";
      GC04_FB13 : "UDT_Conv_G115D_Diagnostics";
      GC04_FB14 : "UDT_Conv_G115D_Diagnostics";
      GC04_FB15 : "UDT_Conv_G115D_Diagnostics";
      GC04_FB16 : "UDT_Conv_G115D_Diagnostics";
      GC04_FB17 : "UDT_Conv_G115D_Diagnostics";
      GC04_FB18 : "UDT_Conv_G115D_Diagnostics";
      GC04_FB19 : "UDT_Conv_G115D_Diagnostics";
      GC04_RC20 : "UDT_Conv_MultiControl_Diagnostics";
      GC04_RC21_Track : "UDT_Track_Statistics";
      GC04_RC21 : "UDT_Conv_Dual_G115D_Diagnostics";
      GC05_RC01 : "UDT_Conv_MultiControl_Diagnostics";
      GC05_RC02 : "UDT_Conv_MultiControl_Diagnostics";
      GC05_RC03 : "UDT_Conv_MultiControl_Diagnostics";
      GC05_RC10 : "UDT_Conv_MultiControl_Diagnostics";
      GC05_FB04 : "UDT_Conv_G115D_Diagnostics";
      GC05_FB05 : "UDT_Conv_G115D_Diagnostics";
      GC05_RC06 : "UDT_Conv_MultiControl_Diagnostics";
      GC05_RC07 : "UDT_Conv_G115D_Diagnostics";
      GC06_RC01 : "UDT_Conv_MultiControl_Diagnostics";
      GC06_FB02 : "UDT_Conv_G115D_Diagnostics";
      GC06_FB03 : "UDT_Conv_G115D_Diagnostics";
      GC06_RC04 : "UDT_Conv_Triple_G115D_Diagnostics";
      GC06_FB05 : "UDT_Conv_G115D_Diagnostics";
      GC06_FB06 : "UDT_Conv_G115D_Diagnostics";
      GC06_FB07 : "UDT_Conv_G115D_Diagnostics";
      GC06_SK08 : "UDT_Conv_G115D_Diagnostics";
      GC07_CH01 : "UDT_Chute_Statistics";
      GC07_FB01 : "UDT_Conv_G115D_Diagnostics";
      GC07_RC02 : "UDT_Conv_Dual_G115D_Diagnostics";
      GC07_RC03 : "UDT_Conv_MultiControl_Diagnostics";
      GC07_RC04 : "UDT_Conv_MultiControl_Diagnostics";
      GC07_RC05 : "UDT_Conv_MultiControl_Diagnostics";
      GC07_RC06 : "UDT_Conv_MultiControl_Diagnostics";
      GC07_RC10 : "UDT_Conv_MultiControl_Diagnostics";
      GC07_RC07 : "UDT_Conv_MultiControl_Diagnostics";
      GC07_RC08 : "UDT_Conv_MultiControl_Diagnostics";
      GC07_RC11 : "UDT_Conv_MultiControl_Diagnostics";
      GC07_CH02 : "UDT_Divert_Statistics";
      GC07_FB09 : "UDT_Conv_G115D_Diagnostics";
   END_VAR


BEGIN

END_DATA_BLOCK

FUNCTION_BLOCK "FB_SINA_SPEED_TEL1"
TITLE = 'Speed Control with SINAMICS and S7'
{ S7_Optimized_Access := 'TRUE' }
AUTHOR : DRVDPS7
FAMILY : DRIVES
NAME : SINA_SPD
VERSION : 5.1
//Copyright (C) Siemens AG 2012. All Rights Reserved. Confidential
//--------------------------------------------------------------------------------------
//SINA_SPEED: Drehzahlregelung mit dem Antriebsbaustein SINAMICS S120/G120 <-> S7-1200
//------------------------------------------------------------------------------------- Ersteller: Siemens AG Erlangen A&D MC PM   Datum:  07.07.10        Vers.:2.1
//Änderung:  J.B. Typical Team                       07.12.12              2.2
//    Umsetzung in SCL / TIA
//Änderung:  J.B. Typical Team                       29.04.13              2.3
//    1. "Q" an den AusgÃ¤nge entfernen
//    2. Neuer Ausgang PwrInhibit
//Änderung:  J.B. Typical Team                       28.06.13              2.4
//    Ã„nderung HW-Zugriff Ã¼ber LOG2MOD
//
//Änderung:  J.B. Typical Team                       18.07.13              2.5
//    Ã„nderung HW-Zugriff Ã¼ber zwei HW-EingÃ¤nge
//
//Änderung:  J.B. Typical Team                       17.07.14              3.0
//    Optimmierung
//
//Änderung:  J.B. Typical Team                       30.07.14              4.0
//    Festlegung auf einheitlicher neuer Version 4.0
//
//Änderung:  P.Z. Typical Team                       03.12.15              4.1
//    Schnittstelle an Programmierleitfadeb TIA-Potal angepasst
//    zusÃ¤tzlicher Eingang "ConfigAxis" fÃ¼r STW-Bits
//
//Änderung:  G.F. Typical Team                       01.03.16              4.2
//    Sollwert auf INT - Grenzen begrenzt
//Änderung:  F.G. Typical Team                       13.09.16              4.3
//    Ausgabewerte am Ausgang "Status" angepasst
//
//Änderung:  G.F. Typical Team                       11.01.17              5.0
//    - Festlegung auf einheitlicher neuer Version 5.0
//
//Änderung:  G.F. Typical Team                       03.05.18              5.1
//    - Alle Bits des Eingang ConfigAxis auf STW1 aufgelegt
//
//Bibliothek V7
//Funktion: Drehzahlregelung mit dem Antriebsbaustein SINAMICS S120/G120 <-> S7-1200
//********************************************************************************************************************************************************
//************************************************************************FB283***************************************************************************
//********************************************************************************************************************************************************
   VAR_INPUT
      EnableAxis : Bool;   // 0-->1; 1 = Enable the drive (OFF2 / OFF 3 are 1 in default status) (OFF1 = 0-->1)
      AckError : Bool;   // 1 = Acknowledge drive error
      SpeedSetpoint : Int;   // Speed standardises with the standardisation factor
      RefSpeed : Int;   // Standardisation factor of speed
      Acceleration : Int;   // Ramp up
      Deceleration : Int;   // Ramp down
      RefRampTime : Int;   // Ramp time reference for ref speed
      ConfigAxis : Word := 16#003F;   // binary programmed input to control all functions in the telegram without its own function block input
   END_VAR

   VAR_OUTPUT
      AxisEnabled : Bool;   // 1 = Drive is enabled
      Lockout : Bool;   // 1 = Drive lockout active
      Fault : Bool;   // 1 = Fault
      Alarm : Bool;   // 1 = Alarm
      ActualSpeed : Int;   // Actual in [U/min]
      FaultCode : Word;
      AlarmCode : Word;
   END_VAR

   VAR_IN_OUT
      io_HW_Interface : "UDT_G115D_HW_Interface";
   END_VAR

   VAR CONSTANT
      C_MIN_SCALE : Real := -32768.0;
      C_MAX_SCALE : Real := 32767.0;
   END_VAR


BEGIN
	//=============================================================================
	//SIEMENS AG
	//(c)Copyright 2017 All Rights Reserved
	//-----------------------------------------------------------------------------
	// Library: DriveLib - UDT Updated Version
	// Function: Speed control with SINAMICS using UDT interface
	//=============================================================================

	// Evaluate drive status from UDT bits
	#AxisEnabled := #io_HW_Interface.Input.ZSW1_Bit02_Enabled;     // Bit 2: Operation enabled
	#Fault := #io_HW_Interface.Input.ZSW1_Bit03_Fault OR #io_HW_Interface.Input.ZSW_G115D_Bit08_PowerOff;             // Bit 3: Fault
	#Alarm := #io_HW_Interface.Input.ZSW1_Bit07_Alarm;             // Bit 7: Alarm
	#Lockout := #io_HW_Interface.Input.ZSW1_Bit06_Inhibit;         // Bit 6: Switching on inhibited
	#FaultCode := #io_HW_Interface.Input.FaultCode;
	#AlarmCode := #io_HW_Interface.Input.AlarmCode;

	// Calculate actual velocity from NIST_A
	IF #RefSpeed <> 0 THEN
	    #ActualSpeed := REAL_TO_INT(INT_TO_REAL(#io_HW_Interface.Input.NIST_A) / 16384.0 * INT_TO_REAL(#RefSpeed));
	ELSE
	    #ActualSpeed := 0;
	END_IF;

	// Build control word using UDT unpacked bits
	// STW1 bit mapping using UDT variables instead of slice access

	// Bit 0: ON/OFF1 (EnableAxis)
	#io_HW_Interface.Output.STW1_Bit00_On := #EnableAxis;

	// Bit 1: OFF2 (from ConfigAxis bit 0, inverted logic: 1=active/no OFF2)
	#io_HW_Interface.Output.STW1_Bit01_Off2 := #ConfigAxis.%X0;

	// Bit 2: OFF3 (from ConfigAxis bit 1, inverted logic: 1=active/no OFF3)
	#io_HW_Interface.Output.STW1_Bit02_Off3 := #ConfigAxis.%X1;

	// Bit 3: Operation enable (from ConfigAxis bit 2)
	#io_HW_Interface.Output.STW1_Bit03_Enable := #ConfigAxis.%X2;

	// Bit 4: Ramp enable (from ConfigAxis bit 3)
	#io_HW_Interface.Output.STW1_Bit04_RampEnable := #ConfigAxis.%X3;

	// Bit 5: Ramp continue (from ConfigAxis bit 4)
	#io_HW_Interface.Output.STW1_Bit05_RampContinue := #ConfigAxis.%X4;

	// Bit 6: Setpoint enable (from ConfigAxis bit 5)
	#io_HW_Interface.Output.STW1_Bit06_SetEnable := #ConfigAxis.%X5;

	// Bit 7: Acknowledge fault
	#io_HW_Interface.Output.STW1_Bit07_Ack := #AckError;

	// Bit 8: Reserved (from ConfigAxis bit 10)
	#io_HW_Interface.Output.STW1_Bit08_Reserved := #ConfigAxis.%X10;

	// Bit 9: Reserved (from ConfigAxis bit 11)
	#io_HW_Interface.Output.STW1_Bit09_Reserved := #ConfigAxis.%X11;

	// Bit 10: Control by PLC (must be TRUE)
	#io_HW_Interface.Output.STW1_Bit10_PLC := TRUE;

	// Bit 11: Reverse direction (from ConfigAxis bit 6)
	#io_HW_Interface.Output.STW1_Bit11_Reverse := #ConfigAxis.%X6;

	// Bit 12: Reserved (from ConfigAxis bit 7)
	#io_HW_Interface.Output.STW1_Bit12_Reserved := #ConfigAxis.%X7;

	// Bit 13: MOP up (from ConfigAxis bit 8)
	#io_HW_Interface.Output.STW1_Bit13_MOP_Up := #ConfigAxis.%X8;

	// Bit 14: MOP down (from ConfigAxis bit 9)
	#io_HW_Interface.Output.STW1_Bit14_MOP_Down := #ConfigAxis.%X9;

	// Bit 15: Reserved (from ConfigAxis bit 12)
	#io_HW_Interface.Output.STW1_Bit15_Reserved := #ConfigAxis.%X12;

	// Calculate velocity setpoint
	IF #RefSpeed <> 0.0 THEN
	    #io_HW_Interface.Output.NSOLL_A := REAL_TO_INT(
	                                                   LIMIT_REAL(MN := #C_MIN_SCALE,
	                                                              IN := INT_TO_REAL(#SpeedSetpoint) * (16384.0 / INT_TO_REAL(#RefSpeed)),
	                                                              MX := #C_MAX_SCALE));
	ELSE
	    #io_HW_Interface.Output.NSOLL_A := 0;
	END_IF;

	#io_HW_Interface.Output.RampUpScaling := REAL_TO_INT(
	                                                     LIMIT_REAL(MN := 0,
	                                                                IN := INT_TO_REAL(#RefSpeed) / INT_TO_REAL(#Acceleration) * 1000 / INT_TO_REAL(#RefRampTime) * 16384.0,
	                                                                MX := #C_MAX_SCALE));
	#io_HW_Interface.Output.RampDownScaling := REAL_TO_INT(
	                                                       LIMIT_REAL(MN := 0,
	                                                                  IN := INT_TO_REAL(#RefSpeed) / INT_TO_REAL(#Deceleration) * 1000 / INT_TO_REAL(#RefRampTime) * 16384.0,
	                                                                  MX := #C_MAX_SCALE));

END_FUNCTION_BLOCK

FUNCTION "FC_IFM_VFD_G115D_In" : Void
{ S7_Optimized_Access := 'TRUE' }
VERSION : 0.1
   VAR_INPUT
      i_Telegram_HW_ID : HW_SUBMODULE;
      i_Additional_HW_ID : HW_SUBMODULE;
   END_VAR

   VAR_OUTPUT
      o_Telegram_Start_Address : Int;
      o_ActualValue_Start_Address : Int;
      o_Data : "UDT_G115D_HW_Input";
   END_VAR

   VAR_TEMP
      t_ZSW1_Word : Word;
      t_ZSW_G115D_Word : Word;
      t_ZSW2_G115D_Word : Word;
      t_Value_Byte : Byte;
      t_Ret_Val_Int : Int;
      t_HW_RD_Inf_Rec_I_Address : UDInt;
      t_HW_RD_Inf_Rec_I_Len : UInt;
      t_HW_WR_Inf_Rec_O_Address : UDInt;
      t_HW_WR_Inf_Rec_O_Len : UInt;
      t_Word_Scale_Data : Word;
   END_VAR

   VAR CONSTANT
      C_REF_VOLTAGE : Int := 1000;   // [V]
      C_REF_CURRENT : Int := 10;   // [A]
      C_REF_TORQUE : Int := 100;   // [Nm]
      C_REF_POWER : Int := 31420;   // [W]
      C_REF_TEMP : Int := 100;   // [°C]
   END_VAR


BEGIN
	REGION Telegram Module
	    #t_ZSW1_Word := 0;

	    #t_Ret_Val_Int := RD_ADDR(LADDR := #i_Telegram_HW_ID,
	                              PIADDR => #t_HW_RD_Inf_Rec_I_Address,
	                              PICount => #t_HW_RD_Inf_Rec_I_Len,
	                              PQADDR => #t_HW_WR_Inf_Rec_O_Address,
	                              PQCount => #t_HW_WR_Inf_Rec_O_Len);

	    #o_Telegram_Start_Address := UDINT_TO_INT(#t_HW_RD_Inf_Rec_I_Address);

	    IF #t_Ret_Val_Int = 0 AND #t_HW_RD_Inf_Rec_I_Len = 4 THEN
	        #t_ZSW1_Word := PEEK_WORD(area := 16#81, // Input area
	                                  dbNumber := 0,
	                                  byteOffset := UDINT_TO_DINT(#t_HW_RD_Inf_Rec_I_Address));

	        #o_Data.NIST_A := PEEK_WORD(area := 16#81, // Input area
	                                    dbNumber := 0,
	                                    byteOffset := UDINT_TO_DINT(#t_HW_RD_Inf_Rec_I_Address) + 2);
	    ELSE
	        #o_Data.NIST_A := 0;
	    END_IF;
	    #o_Data.ZSW1_Bit00_ReadyOn := #t_ZSW1_Word.%X0;
	    #o_Data.ZSW1_Bit01_Ready := #t_ZSW1_Word.%X1;
	    #o_Data.ZSW1_Bit02_Enabled := #t_ZSW1_Word.%X2;
	    #o_Data.ZSW1_Bit03_Fault := #t_ZSW1_Word.%X3;
	    #o_Data.ZSW1_Bit04_NoCoastActive := #t_ZSW1_Word.%X4;
	    #o_Data.ZSW1_Bit05_NoQuickStopActive := #t_ZSW1_Word.%X5;
	    #o_Data.ZSW1_Bit06_Inhibit := #t_ZSW1_Word.%X6;
	    #o_Data.ZSW1_Bit07_Alarm := #t_ZSW1_Word.%X7;
	    #o_Data.ZSW1_Bit08_DeviationOK := #t_ZSW1_Word.%X8;
	    #o_Data.ZSW1_Bit09_ControlQuest := #t_ZSW1_Word.%X9;
	    #o_Data.ZSW1_Bit10_OverSpeed := #t_ZSW1_Word.%X10;
	    #o_Data.ZSW1_Bit11_Limit := #t_ZSW1_Word.%X11;
	    #o_Data.ZSW1_Bit12_Brake := #t_ZSW1_Word.%X12;
	    #o_Data.ZSW1_Bit13_MotorTempOK := #t_ZSW1_Word.%X13;
	    #o_Data.ZSW1_Bit14_Direction_CW := #t_ZSW1_Word.%X14;
	    #o_Data.ZSW1_Bit15_VFDTempOK := #t_ZSW1_Word.%X15;
	END_REGION

	REGION Actual Value Module
	    #t_ZSW_G115D_Word := 0;
	    #t_ZSW2_G115D_Word := 0;

	    #t_Ret_Val_Int := RD_ADDR(LADDR := #i_Additional_HW_ID,
	                              PIADDR => #t_HW_RD_Inf_Rec_I_Address,
	                              PICount => #t_HW_RD_Inf_Rec_I_Len,
	                              PQADDR => #t_HW_WR_Inf_Rec_O_Address,
	                              PQCount => #t_HW_WR_Inf_Rec_O_Len);

	    #o_ActualValue_Start_Address := UDINT_TO_INT(#t_HW_RD_Inf_Rec_I_Address);

	    IF #t_Ret_Val_Int = 0 AND #t_HW_RD_Inf_Rec_I_Len = 20 THEN
	        #t_ZSW_G115D_Word := PEEK_WORD(area := 16#81, // Input area
	                                       dbNumber := 0,
	                                       byteOffset := UDINT_TO_DINT(#t_HW_RD_Inf_Rec_I_Address));

	        #o_Data.FaultCode := PEEK_WORD(area := 16#81, // Input area
	                                       dbNumber := 0,
	                                       byteOffset := UDINT_TO_DINT(#t_HW_RD_Inf_Rec_I_Address) + 2);

	        #o_Data.AlarmCode := PEEK_WORD(area := 16#81, // Input area
	                                      dbNumber := 0,
	                                      byteOffset := UDINT_TO_DINT(#t_HW_RD_Inf_Rec_I_Address) + 4);

	        #t_Word_Scale_Data := PEEK_WORD(area := 16#81, // Input area
	                                        dbNumber := 0,
	                                        byteOffset := UDINT_TO_DINT(#t_HW_RD_Inf_Rec_I_Address) + 6);

	        #o_Data.DCLinkVoltage := DINT_TO_INT(WORD_TO_DINT(#t_Word_Scale_Data) * #C_REF_VOLTAGE / 16#4000);

	        #t_Word_Scale_Data := PEEK_WORD(area := 16#81, // Input area
	                                        dbNumber := 0,
	                                        byteOffset := UDINT_TO_DINT(#t_HW_RD_Inf_Rec_I_Address) + 8);

	        #o_Data.ActualCurrent := DINT_TO_INT(WORD_TO_DINT(#t_Word_Scale_Data) * #C_REF_CURRENT * 10 / 16#4000);

	        #t_Word_Scale_Data := PEEK_WORD(area := 16#81, // Input area
	                                        dbNumber := 0,
	                                        byteOffset := UDINT_TO_DINT(#t_HW_RD_Inf_Rec_I_Address) + 10);

	        #o_Data.ActivePower := DINT_TO_INT(WORD_TO_DINT(#t_Word_Scale_Data) * #C_REF_POWER / 16#4000);

	        #t_ZSW2_G115D_Word := PEEK_WORD(area := 16#81, // Input area
	                                       dbNumber := 0,
	                                       byteOffset := UDINT_TO_DINT(#t_HW_RD_Inf_Rec_I_Address) + 12);
	    ELSE
	        #o_Data.FaultCode := 0;
	        #o_Data.AlarmCode := 0;
	        #o_Data.DCLinkVoltage := 0;
	        #o_Data.ActualCurrent := 0;
	        #o_Data.ActivePower := 0;
	    END_IF;
	    #o_Data.ZSW_G115D_Bit00_DI0 := #t_ZSW_G115D_Word.%X0;
	    #o_Data.ZSW_G115D_Bit01_DI1 := #t_ZSW_G115D_Word.%X1;
	    #o_Data.ZSW_G115D_Bit02_DI2 := #t_ZSW_G115D_Word.%X2;
	    #o_Data.ZSW_G115D_Bit03_DI3 := #t_ZSW_G115D_Word.%X3;
	    #o_Data.ZSW_G115D_Bit04_DIO24 := #t_ZSW_G115D_Word.%X4;
	    #o_Data.ZSW_G115D_Bit05_DIO25 := #t_ZSW_G115D_Word.%X5;
	    #o_Data.ZSW_G115D_Bit06_STOActive := #t_ZSW_G115D_Word.%X6;
	    #o_Data.ZSW_G115D_Bit07_Reserved := #t_ZSW_G115D_Word.%X7;
	    #o_Data.ZSW_G115D_Bit08_PowerOff := #t_ZSW_G115D_Word.%X8;
	    #o_Data.ZSW_G115D_Bit09_Auto := #t_ZSW_G115D_Word.%X9;
	    #o_Data.ZSW_G115D_Bit10_Manual := #t_ZSW_G115D_Word.%X10;
	    #o_Data.ZSW_G115D_Bit11_Bypass := #t_ZSW_G115D_Word.%X11;
	    #o_Data.ZSW_G115D_Bit12_ContMotion := #t_ZSW_G115D_Word.%X12;
	    #o_Data.ZSW_G115D_Bit13_JogLeft := #t_ZSW_G115D_Word.%X13;
	    #o_Data.ZSW_G115D_Bit14_JogRight := #t_ZSW_G115D_Word.%X14;
	    #o_Data.ZSW_G115D_Bit15_Reserved := #t_ZSW_G115D_Word.%X15;

	    #o_Data.ZSW2_G115D_Bit00_Memory_Card_In := #t_ZSW2_G115D_Word.%X0;
	    #o_Data.ZSW2_G115D_Bit01_Memory_Card_Active := #t_ZSW2_G115D_Word.%X1;
	    #o_Data.ZSW2_G115D_Bit02_Memory_Card_Siemens := #t_ZSW2_G115D_Word.%X2;
	    #o_Data.ZSW2_G115D_Bit03_Memory_Card_USB := #t_ZSW2_G115D_Word.%X3;
	    #o_Data.ZSW2_G115D_Bit04_Reserved := #t_ZSW2_G115D_Word.%X4;
	    #o_Data.ZSW2_G115D_Bit05_Reserved := #t_ZSW2_G115D_Word.%X5;
	    #o_Data.ZSW2_G115D_Bit06_Reserved := #t_ZSW2_G115D_Word.%X6;
	    #o_Data.ZSW2_G115D_Bit07_Reserved := #t_ZSW2_G115D_Word.%X7;
	    #o_Data.ZSW2_G115D_Bit08_Reserved := #t_ZSW2_G115D_Word.%X8;
	    #o_Data.ZSW2_G115D_Bit09_Reserved := #t_ZSW2_G115D_Word.%X9;
	    #o_Data.ZSW2_G115D_Bit10_Reserved := #t_ZSW2_G115D_Word.%X10;
	    #o_Data.ZSW2_G115D_Bit11_Reserved := #t_ZSW2_G115D_Word.%X11;
	    #o_Data.ZSW2_G115D_Bit12_Reserved := #t_ZSW2_G115D_Word.%X12;
	    #o_Data.ZSW2_G115D_Bit13_Reserved := #t_ZSW2_G115D_Word.%X13;
	    #o_Data.ZSW2_G115D_Bit14_Reserved := #t_ZSW2_G115D_Word.%X14;
	    #o_Data.ZSW2_G115D_Bit15_Reserved := #t_ZSW2_G115D_Word.%X15;
	END_REGION
END_FUNCTION

FUNCTION "FC_IFM_VFD_G115D_Out" : Void
{ S7_Optimized_Access := 'TRUE' }
VERSION : 0.1
   VAR_INPUT
      i_Telegram_HW_ID : HW_SUBMODULE;
      i_Additional_HW_ID : HW_SUBMODULE;
      i_Data : "UDT_G115D_HW_Output";
   END_VAR

   VAR_OUTPUT
      o_Telegram_Start_Address : Int;
      o_ActualValue_Start_Address : Int;
   END_VAR

   VAR_TEMP
      t_STW1_Word : Word;
      t_STW_G115D_Word : Word;
      t_Value_Byte : Byte;
      t_Ret_Val_Int : Int;
      t_HW_RD_Inf_Rec_I_Address : UDInt;
      t_HW_RD_Inf_Rec_I_Len : UInt;
      t_HW_WR_Inf_Rec_O_Address : UDInt;
      t_HW_WR_Inf_Rec_O_Len : UInt;
   END_VAR


BEGIN
	REGION Telegram Module
	    #t_STW1_Word := 0;

	    #t_Ret_Val_Int := RD_ADDR(LADDR := #i_Telegram_HW_ID,
	                              PIADDR => #t_HW_RD_Inf_Rec_I_Address,
	                              PICount => #t_HW_RD_Inf_Rec_I_Len,
	                              PQADDR => #t_HW_WR_Inf_Rec_O_Address,
	                              PQCount => #t_HW_WR_Inf_Rec_O_Len);

	    #o_Telegram_Start_Address := UDINT_TO_INT(#t_HW_WR_Inf_Rec_O_Address);

	    #t_STW1_Word.%X0 := #i_Data.STW1_Bit00_On;
	    #t_STW1_Word.%X1 := #i_Data.STW1_Bit01_Off2;
	    #t_STW1_Word.%X2 := #i_Data.STW1_Bit02_Off3;
	    #t_STW1_Word.%X3 := #i_Data.STW1_Bit03_Enable;
	    #t_STW1_Word.%X4 := #i_Data.STW1_Bit04_RampEnable;
	    #t_STW1_Word.%X5 := #i_Data.STW1_Bit05_RampContinue;
	    #t_STW1_Word.%X6 := #i_Data.STW1_Bit06_SetEnable;
	    #t_STW1_Word.%X7 := #i_Data.STW1_Bit07_Ack;
	    #t_STW1_Word.%X8 := #i_Data.STW1_Bit08_Reserved;
	    #t_STW1_Word.%X9 := #i_Data.STW1_Bit09_Reserved;
	    #t_STW1_Word.%X10 := #i_Data.STW1_Bit10_PLC;
	    #t_STW1_Word.%X11 := #i_Data.STW1_Bit11_Reverse;
	    #t_STW1_Word.%X12 := #i_Data.STW1_Bit12_Reserved;
	    #t_STW1_Word.%X13 := #i_Data.STW1_Bit13_MOP_Up;
	    #t_STW1_Word.%X14 := #i_Data.STW1_Bit14_MOP_Down;
	    #t_STW1_Word.%X15 := #i_Data.STW1_Bit15_Reserved;
	    //#t_STW1_Word := SWAP_WORD(#t_STW1_Word);

	    IF #t_Ret_Val_Int = 0 AND #t_HW_WR_Inf_Rec_O_Len = 4 THEN
	        POKE(area       := 16#82, // Output Area,
	             dbNumber   := 0,
	             byteOffset := UDINT_TO_DINT(#t_HW_WR_Inf_Rec_O_Address),
	             value      := #t_STW1_Word);

	        POKE(area       := 16#82, // Output Area,
	             dbNumber   := 0,
	             byteOffset := UDINT_TO_DINT(#t_HW_WR_Inf_Rec_O_Address) + 2,
	             value      := #i_Data.NSOLL_A);
	    END_IF;
	END_REGION

	REGION Actual Value Module
	    #t_STW_G115D_Word := 0;

	    #t_Ret_Val_Int := RD_ADDR(LADDR := #i_Additional_HW_ID,
	                              PIADDR => #t_HW_RD_Inf_Rec_I_Address,
	                              PICount => #t_HW_RD_Inf_Rec_I_Len,
	                              PQADDR => #t_HW_WR_Inf_Rec_O_Address,
	                              PQCount => #t_HW_WR_Inf_Rec_O_Len);

	    #o_ActualValue_Start_Address := UDINT_TO_INT(#t_HW_WR_Inf_Rec_O_Address);

	    #t_STW_G115D_Word.%X0 := #i_Data.STW_G115D_Bit00_DO24;
	    #t_STW_G115D_Word.%X1 := #i_Data.STW_G115D_Bit01_DO25;
	    #t_STW_G115D_Word.%X2 := #i_Data.STW_G115D_Bit02_Disable_StopSlow_Sensor;
	    #t_STW_G115D_Word.%X3 := #i_Data.STW_G115D_Bit03_Reserved;
	    #t_STW_G115D_Word.%X4 := #i_Data.STW_G115D_Bit04_Reserved;
	    #t_STW_G115D_Word.%X5 := #i_Data.STW_G115D_Bit05_Reserved;
	    #t_STW_G115D_Word.%X6 := #i_Data.STW_G115D_Bit06_Reserved;
	    #t_STW_G115D_Word.%X7 := #i_Data.STW_G115D_Bit07_Reserved;
	    #t_STW_G115D_Word.%X8 := #i_Data.STW_G115D_Bit08_Reserved;
	    #t_STW_G115D_Word.%X9 := #i_Data.STW_G115D_Bit09_Reserved;
	    #t_STW_G115D_Word.%X10 := #i_Data.STW_G115D_Bit10_Reserved;
	    #t_STW_G115D_Word.%X11 := #i_Data.STW_G115D_Bit11_Reserved;
	    #t_STW_G115D_Word.%X12 := #i_Data.STW_G115D_Bit12_Reserved;
	    #t_STW_G115D_Word.%X13 := #i_Data.STW_G115D_Bit13_Reserved;
	    #t_STW_G115D_Word.%X14 := #i_Data.STW_G115D_Bit14_Reserved;
	    #t_STW_G115D_Word.%X15 := #i_Data.STW_G115D_Bit15_Reserved;
	    //#t_STW_G115D_Word := SWAP_WORD(#t_STW_G115D_Word);

	    IF #t_Ret_Val_Int = 0 AND #t_HW_WR_Inf_Rec_O_Len = 20 THEN
	        POKE(area       := 16#82, // Output Area,
	             dbNumber   := 0,
	             byteOffset := UDINT_TO_DINT(#t_HW_WR_Inf_Rec_O_Address),
	             value      := #t_STW_G115D_Word);

	        POKE(area       := 16#82, // Output Area,
	             dbNumber   := 0,
	             byteOffset := UDINT_TO_DINT(#t_HW_WR_Inf_Rec_O_Address) + 2,
	             value      := #i_Data.RampUpScaling);

	        POKE(area       := 16#82, // Output Area,
	             dbNumber   := 0,
	             byteOffset := UDINT_TO_DINT(#t_HW_WR_Inf_Rec_O_Address) + 4,
	             value      := #i_Data.RampDownScaling);
	    END_IF;
	END_REGION
END_FUNCTION

FUNCTION "FC_IFM_VFD_S210_Out" : Void
{ S7_Optimized_Access := 'TRUE' }
VERSION : 0.1
   VAR_INPUT
      i_Telegram_HW_ID : HW_SUBMODULE;
      i_Data : "UDT_S210_HW_Output";
   END_VAR

   VAR_OUTPUT
      o_Telegram_Start_Address : Int;
      o_ActualValue_Start_Address : Int;
   END_VAR

   VAR_TEMP
      t_STW1_Word : Word;
      t_POS_STW1_Word : Word;
      t_POS_STW2_Word : Word;
      t_STW2_Word : Word;
      t_Value_Byte : Byte;
      t_Ret_Val_Int : Int;
      t_HW_RD_Inf_Rec_I_Address : UDInt;
      t_HW_RD_Inf_Rec_I_Len : UInt;
      t_HW_WR_Inf_Rec_O_Address : UDInt;
      t_HW_WR_Inf_Rec_O_Len : UInt;
   END_VAR


BEGIN
	REGION Telegram Module
	    #t_STW1_Word := 0;
	    #t_POS_STW1_Word := 0;
	    #t_POS_STW2_Word := 0;
	    #t_STW2_Word := 0;

	    #t_Ret_Val_Int := RD_ADDR(LADDR := #i_Telegram_HW_ID,
	                              PIADDR => #t_HW_RD_Inf_Rec_I_Address,
	                              PICount => #t_HW_RD_Inf_Rec_I_Len,
	                              PQADDR => #t_HW_WR_Inf_Rec_O_Address,
	                              PQCount => #t_HW_WR_Inf_Rec_O_Len);

	    #o_Telegram_Start_Address := UDINT_TO_INT(#t_HW_WR_Inf_Rec_O_Address);

	    // Pack STW1 bits
	    #t_STW1_Word.%X0 := #i_Data.STW1_Bit00_On;
	    #t_STW1_Word.%X1 := #i_Data.STW1_Bit01_Off2;
	    #t_STW1_Word.%X2 := #i_Data.STW1_Bit02_Off3;
	    #t_STW1_Word.%X3 := #i_Data.STW1_Bit03_Enable;
	    #t_STW1_Word.%X4 := #i_Data.STW1_Bit04_NotRejectTask;
	    #t_STW1_Word.%X5 := #i_Data.STW1_Bit05_NoIntermediateStop;
	    #t_STW1_Word.%X6 := #i_Data.STW1_Bit06_ActivateTask;
	    #t_STW1_Word.%X7 := #i_Data.STW1_Bit07_Ack;
	    #t_STW1_Word.%X8 := #i_Data.STW1_Bit08_Jog1;
	    #t_STW1_Word.%X9 := #i_Data.STW1_Bit09_Jog2;
	    #t_STW1_Word.%X10 := #i_Data.STW1_Bit10_PLC;
	    #t_STW1_Word.%X11 := #i_Data.STW1_Bit11_StartHoming;
	    #t_STW1_Word.%X12 := #i_Data.STW1_Bit12_Reserved;
	    #t_STW1_Word.%X13 := #i_Data.STW1_Bit13_ExtBlockChange;
	    #t_STW1_Word.%X14 := #i_Data.STW1_Bit14_Reserved;
	    #t_STW1_Word.%X15 := #i_Data.STW1_Bit15_Reserved;

	    // Pack POS_STW1 bits
	    #t_POS_STW1_Word.%X0 := #i_Data.POS_STW1_Bit00_Traversing0;
	    #t_POS_STW1_Word.%X1 := #i_Data.POS_STW1_Bit01_Traversing1;
	    #t_POS_STW1_Word.%X2 := #i_Data.POS_STW1_Bit02_Traversing2;
	    #t_POS_STW1_Word.%X3 := #i_Data.POS_STW1_Bit03_Traversing3;
	    #t_POS_STW1_Word.%X4 := #i_Data.POS_STW1_Bit04_Traversing4;
	    #t_POS_STW1_Word.%X5 := #i_Data.POS_STW1_Bit05_Traversing5;
	    #t_POS_STW1_Word.%X6 := #i_Data.POS_STW1_Bit06_Reserved;
	    #t_POS_STW1_Word.%X7 := #i_Data.POS_STW1_Bit07_ReleaseBrake;
	    #t_POS_STW1_Word.%X8 := #i_Data.POS_STW1_Bit08_Absolute;
	    #t_POS_STW1_Word.%X9 := #i_Data.POS_STW1_Bit09_DirPos;
	    #t_POS_STW1_Word.%X10 := #i_Data.POS_STW1_Bit10_DirNeg;
	    #t_POS_STW1_Word.%X11 := #i_Data.POS_STW1_Bit11_Reserved;
	    #t_POS_STW1_Word.%X12 := #i_Data.POS_STW1_Bit12_Continuous;
	    #t_POS_STW1_Word.%X13 := #i_Data.POS_STW1_Bit13_Reserved;
	    #t_POS_STW1_Word.%X14 := #i_Data.POS_STW1_Bit14_SetupOrPositioning;
	    #t_POS_STW1_Word.%X15 := #i_Data.POS_STW1_Bit15_ActivateMDI;

	    // Pack POS_STW2 bits
	    #t_POS_STW2_Word.%X0 := #i_Data.POS_STW2_Bit00_ActivateFollowUp;
	    #t_POS_STW2_Word.%X1 := #i_Data.POS_STW2_Bit01_SetRefPoint;
	    #t_POS_STW2_Word.%X2 := #i_Data.POS_STW2_Bit02_RefCam;
	    #t_POS_STW2_Word.%X3 := #i_Data.POS_STW2_Bit03_AdjustEncoder;
	    #t_POS_STW2_Word.%X4 := #i_Data.POS_STW2_Bit04_Reserved;
	    #t_POS_STW2_Word.%X5 := #i_Data.POS_STW2_Bit05_JogIncrementalOrVelocity;
	    #t_POS_STW2_Word.%X6 := #i_Data.POS_STW2_Bit06_Reserved;
	    #t_POS_STW2_Word.%X7 := #i_Data.POS_STW2_Bit07_Reserved;
	    #t_POS_STW2_Word.%X8 := #i_Data.POS_STW2_Bit08_RefType;
	    #t_POS_STW2_Word.%X9 := #i_Data.POS_STW2_Bit09_RefNegDir;
	    #t_POS_STW2_Word.%X10 := #i_Data.POS_STW2_Bit10_MeasProbe2;
	    #t_POS_STW2_Word.%X11 := #i_Data.POS_STW2_Bit11_MeasProbeEdge;
	    #t_POS_STW2_Word.%X12 := #i_Data.POS_STW2_Bit12_Reserved;
	    #t_POS_STW2_Word.%X13 := #i_Data.POS_STW2_Bit13_Reserved;
	    #t_POS_STW2_Word.%X14 := #i_Data.POS_STW2_Bit14_SWLimit;
	    #t_POS_STW2_Word.%X15 := #i_Data.POS_STW2_Bit15_StopCam;

	    // Pack STW2 bits
	    #t_STW2_Word.%X0 := #i_Data.STW2_Bit00_Reserved;
	    #t_STW2_Word.%X1 := #i_Data.STW2_Bit01_Reserved;
	    #t_STW2_Word.%X2 := #i_Data.STW2_Bit02_Reserved;
	    #t_STW2_Word.%X3 := #i_Data.STW2_Bit03_Reserved;
	    #t_STW2_Word.%X4 := #i_Data.STW2_Bit04_Reserved;
	    #t_STW2_Word.%X5 := #i_Data.STW2_Bit05_Reserved;
	    #t_STW2_Word.%X6 := #i_Data.STW2_Bit06_Reserved;
	    #t_STW2_Word.%X7 := #i_Data.STW2_Bit07_Reserved;
	    #t_STW2_Word.%X8 := #i_Data.STW2_Bit08_Reserved;
	    #t_STW2_Word.%X9 := #i_Data.STW2_Bit09_Reserved;
	    #t_STW2_Word.%X10 := #i_Data.STW2_Bit10_Reserved;
	    #t_STW2_Word.%X11 := #i_Data.STW2_Bit11_Reserved;
	    #t_STW2_Word.%X12 := #i_Data.STW2_Bit12_Reserved;
	    #t_STW2_Word.%X13 := #i_Data.STW2_Bit13_Reserved;
	    #t_STW2_Word.%X14 := #i_Data.STW2_Bit14_Reserved;
	    #t_STW2_Word.%X15 := #i_Data.STW2_Bit15_Reserved;

	    IF #t_Ret_Val_Int = 0 AND #t_HW_WR_Inf_Rec_O_Len = 34 THEN
	        // PZD1: STW1
	        POKE(area       := 16#82, // Output Area
	             dbNumber   := 0,
	             byteOffset := UDINT_TO_DINT(#t_HW_WR_Inf_Rec_O_Address),
	             value      := #t_STW1_Word);

	        // PZD2: POS_STW1
	        POKE(area       := 16#82,
	             dbNumber   := 0,
	             byteOffset := UDINT_TO_DINT(#t_HW_WR_Inf_Rec_O_Address) + 2,
	             value      := #t_POS_STW1_Word);

	        // PZD3: POS_STW2
	        POKE(area       := 16#82,
	             dbNumber   := 0,
	             byteOffset := UDINT_TO_DINT(#t_HW_WR_Inf_Rec_O_Address) + 4,
	             value      := #t_POS_STW2_Word);

	        // PZD4: STW2
	        POKE(area       := 16#82,
	             dbNumber   := 0,
	             byteOffset := UDINT_TO_DINT(#t_HW_WR_Inf_Rec_O_Address) + 6,
	             value      := #t_STW2_Word);

	        // PZD5: Override (Int)
	        POKE(area       := 16#82,
	             dbNumber   := 0,
	             byteOffset := UDINT_TO_DINT(#t_HW_WR_Inf_Rec_O_Address) + 8,
	             value      := INT_TO_WORD(#i_Data.Override));

	        // PZD6-7: MDI_TARPOS (Real/Float32)
	        POKE(area       := 16#82,
	             dbNumber   := 0,
	             byteOffset := UDINT_TO_DINT(#t_HW_WR_Inf_Rec_O_Address) + 10,
	             value      := REAL_TO_DWORD(#i_Data.MDI_TARPOS));

	        // PZD8-9: MDI_VELOCITY (Real/Float32)
	        POKE(area       := 16#82,
	             dbNumber   := 0,
	             byteOffset := UDINT_TO_DINT(#t_HW_WR_Inf_Rec_O_Address) + 14,
	             value      := REAL_TO_DWORD(#i_Data.MDI_VELOCITY));

	        // PZD10-11: MDI_ACC (Real/Float32)
	        POKE(area       := 16#82,
	             dbNumber   := 0,
	             byteOffset := UDINT_TO_DINT(#t_HW_WR_Inf_Rec_O_Address) + 18,
	             value      := REAL_TO_DWORD(#i_Data.MDI_ACC));

	        // PZD12-13: MDI_DEC (Real/Float32)
	        POKE(area       := 16#82,
	             dbNumber   := 0,
	             byteOffset := UDINT_TO_DINT(#t_HW_WR_Inf_Rec_O_Address) + 22,
	             value      := REAL_TO_DWORD(#i_Data.MDI_DEC));

	        // PZD14-15: Reserved (Real/Float32)
	        POKE(area       := 16#82,
	             dbNumber   := 0,
	             byteOffset := UDINT_TO_DINT(#t_HW_WR_Inf_Rec_O_Address) + 26,
	             value      := REAL_TO_DWORD(#i_Data.Reserved));

	        // PZD16-17: REF_COORDINATE (Real/Float32)
	        POKE(area       := 16#82,
	             dbNumber   := 0,
	             byteOffset := UDINT_TO_DINT(#t_HW_WR_Inf_Rec_O_Address) + 30,
	             value      := REAL_TO_DWORD(#i_Data.REF_COORDINATE));
	    END_IF;
	END_REGION
END_FUNCTION

FUNCTION "FC_Delay_Off" : Void
{ S7_Optimized_Access := 'TRUE' }
VERSION : 0.1
   VAR_INPUT
      i_CMD_Start : Bool;
      i_CFG_Target : Int;
      i_Cycle_Count : Int;
   END_VAR

   VAR_OUTPUT
      o_Delay_Finish : Bool;
   END_VAR

   VAR_IN_OUT
      io_Setpoint : Int;
   END_VAR


BEGIN
	// Init time value
	IF #i_CMD_Start THEN
	    #io_Setpoint := #i_CFG_Target;
	END_IF;

	// Detect result
	#o_Delay_Finish := #i_CMD_Start OR (NOT #i_CMD_Start AND #io_Setpoint > 0);

	// Count time value
	IF NOT #i_CMD_Start THEN
	    #io_Setpoint := #io_Setpoint - #i_Cycle_Count;
	    IF #io_Setpoint < 0 THEN
	        #io_Setpoint := 0;
	    END_IF;
	END_IF;
END_FUNCTION

FUNCTION "FC_Delay_On" : Void
{ S7_Optimized_Access := 'TRUE' }
VERSION : 0.1
   VAR_INPUT
      i_CMD_Start : Bool;
      i_CFG_Target : Int;
      i_Cycle_Count : Int;
   END_VAR

   VAR_OUTPUT
      o_Delay_Finish : Bool;
   END_VAR

   VAR_IN_OUT
      io_Setpoint : Int;
   END_VAR


BEGIN
	// Init time value
	IF NOT #i_CMD_Start THEN
	    #io_Setpoint := 0;
	END_IF;

	// Detect result
	#o_Delay_Finish := #i_CMD_Start AND #io_Setpoint >= #i_CFG_Target;

	// Count time value
	IF #i_CMD_Start THEN
	    #io_Setpoint := #io_Setpoint + #i_Cycle_Count;
	    IF #io_Setpoint > #i_CFG_Target THEN
	        #io_Setpoint := #i_CFG_Target;
	    END_IF;
	END_IF;
END_FUNCTION

FUNCTION "FC_IFM_VFD_S210_In" : Void
{ S7_Optimized_Access := 'TRUE' }
VERSION : 0.1
   VAR_INPUT
      i_Telegram_HW_ID : HW_SUBMODULE;
      i_Additional_HW_ID : HW_SUBMODULE;
   END_VAR

   VAR_OUTPUT
      o_Telegram_Start_Address : Int;
      o_ActualValue_Start_Address : Int;
      o_Data : "UDT_S210_HW_Input";
   END_VAR

   VAR_TEMP
      t_ZSW1_Word : Word;
      t_POS_ZSW1_Word : Word;
      t_POS_ZSW2_Word : Word;
      t_ZSW2_Word : Word;
      t_ZSW_S210_Word : Word;
      t_Value_Byte : Byte;
      t_Ret_Val_Int : Int;
      t_HW_RD_Inf_Rec_I_Address : UDInt;
      t_HW_RD_Inf_Rec_I_Len : UInt;
      t_HW_WR_Inf_Rec_O_Address : UDInt;
      t_HW_WR_Inf_Rec_O_Len : UInt;
      t_Word_Scale_Data : Word;
   END_VAR

